(* Logix 5000 project; controller R400_500_XLS vendor 1 type 14 code 216 rev 31.11; software revision 31.01 *)

TASK MainTask (continuous, watchdog 500 ms) : MainProgram

MODULES
   Local : vendor 1 type 14 code 216 (5069 0, rev 31.11)
        LabWasher2:6:O.0   // Audible Alarm/Red Status Light/Alarm Signal Relay
        LabWasher2:6:O.1   // Dry Contact For Cycle Completed or External Pure Water valve
        LabWasher2:6:O.2   // Dry contact For Alarm
        LabWasher2:6:O.3   // Interior Light
        LabWasher2:6:O.4   // Transfer Valve (Normally Open Valve)
        LabWasher2:6:O.5   // Cycle Status Pilot Light
        LabWasher2:6:O.6   // Condensate Return CoolDown water valve
        LabWasher2:6:O.7   // Not Used
        LabWasher2:7:O.0   // Load door close pilot valve
        LabWasher2:7:O.1   // Load door open pilot valve
        LabWasher2:7:O.2   // Unload door close pilot valve
        LabWasher2:7:O.3   // Unload door open pilot valve
        LabWasher2:7:O.4   // Pump low speed
        LabWasher2:7:O.5   // Pump high speed
        LabWasher2:7:O.6   // Hot water sump fill valve
        LabWasher2:7:O.7   // Sump drain valve (Normally open valve)
        LabWasher2:8:O.0   // Vapor removal fan / Drying fan
        LabWasher2:8:O.1   // Sump steam valve/ Electrical Heater
        LabWasher2:8:O.2   // Pure water sump/ Tank fill valve
        LabWasher2:8:O.3   // Drain cool down water valve
        LabWasher2:8:O.4   // Cold water sump fill valve
        LabWasher2:8:O.5   // PWT Steam Valve / Electric Heater
        LabWasher2:8:O.6   // Heat recovery tank drian valve
        LabWasher2:8:O.7   // Pure water tank outlet valve
        LabWasher2:9:O.0   // Drying heating elements
        LabWasher2:9:O.2   // Condenser high flow cold water valve
        LabWasher2:9:O.3   // Condenser low flow cold water valve
        LabWasher2:9:O.4   // Chemical pump #1
        LabWasher2:9:O.5   // Chemical pump #2
        LabWasher2:9:O.6   // Chemical pump #3
        LabWasher2:9:O.7   // Chemical pump #4
        LabWasher2:2:I.0   // Chemical Pump 1 level switch
        LabWasher2:2:I.1   // Chemical Pump #2 level switch
        LabWasher2:2:I.2   // Chemical Pump #3 level switch
        LabWasher2:2:I.3   // Chemical Pump #4 level switch
        LabWasher2:2:I.4   // Pure water tank level switch
        LabWasher2:2:I.5   // Pure water tank safety level switch
        LabWasher2:1:I.0   // Motor overload
        LabWasher2:1:I.1   // MCR input
        LabWasher2:1:I.2   // Load door obstruction switch
        LabWasher2:1:I.3   // Load door close
        LabWasher2:1:I.4   // Sump low level switch
        LabWasher2:1:I.5   // Sump low level switch
        LabWasher2:1:I.6   // Sump safety level switch
        LabWasher2:1:I.7   // Shelf switch
        LabWasher2:3:I.0   // Unload door obstruction switch
        LabWasher2:3:I.1   // Unload door close
        LabWasher2:3:I.2   // Door Open button Unload side
        LabWasher2:3:I.3   // Door Close/ Sielnce button Unload Side
      Serial : vendor 1 type 12 code 320 (5069 1, rev 1.11, StandardDataDriven RPI 80 ms)
      LabWasher2 : 1734-AENT (Ethernet 192.168.1.2, rev 3.4, Output RPI 20 ms)
         IO11 : 1734-IB8 (PointIO 1, rev 3.1)
         IO22 : 1734-IB8 (PointIO 2, rev 3.1)
         IO33 : 1734-IR2 (PointIO 4, rev 3.1, Input RPI 80 ms)
         IO77 : 1734-IR2 (PointIO 5, rev 3.1, Input RPI 80 ms)
         IO66 : 1734-IB8 (PointIO 3, rev 3.1)
         IO99 : 1734-OB8 (PointIO 9, rev 3.1)
         IO88 : 1734-OB8 (PointIO 8, rev 3.1)
         IO44 : 1734-OB8 (PointIO 6, rev 3.1)
         IO55 : 1734-OB8 (PointIO 7, rev 3.1)
      LabWasher : 1734-AENT (Ethernet 192.168.1.4, rev 3.4, Output RPI 20 ms)   // Chamber inputs/outputs remote module
         IO2 : 1734-IB8 (PointIO 2, rev 3.1, Input RPI 20 ms)   // Digital inputs
              LabWasher:2:I.Data.0   // Chemical Pump #1 level switch
              LabWasher:2:I.Data.1   // Chemical Pump #2 level switch
              LabWasher:2:I.Data.2   // Chemical Pump #3 level switch
              LabWasher:2:I.Data.3   // Chemical Pump #4 level switch
              LabWasher:2:I.Data.4   // Pure water tank level switch
              LabWasher:2:I.Data.5   // Pure water tank safety level switch
              LabWasher:2:I.Data.6   // Pure Water Filling Authorization Signal
         IO3 : 1734-IR2 (PointIO 4, rev 3.1, Input RPI 80 ms)   // Analog input
              LabWasher:4:I.Ch0Data   // Sump RTD
              LabWasher:4:I.Ch1Data   // Drying RTD
              LabWasher:4:I.Ch0Fault   // Sump RTD channel Fault bit
              LabWasher:4:I.Ch1Fault   // Dry RTD channel Fault bit
         IO7 : 1734-IR2 (PointIO 5, rev 3.1, Input RPI 80 ms)   // RTD inputs
              LabWasher:5:I.Ch0Data   // Pure Water Tank RTD
              LabWasher:5:I.Ch1Data   // Not Used
              LabWasher:5:I.Ch0Fault   // Pure Water Tank RTD channel Fault bit
         IO10 : 1734-IE4C (PointIO 10, rev 3.1, Input RPI 80 ms)   // Analog inputs
              LabWasher:10:I.Ch0Data   // Chemical water conductivity
              LabWasher:10:I.Ch1Data   // Final rinse water conductivity
              LabWasher:10:I.Ch2Data   // Recirculation pump pressure
              LabWasher:10:I.Ch3Data   // Not Used
              LabWasher:10:I.Ch0Fault   // Chemical conductivity channel Fault bit
              LabWasher:10:I.Ch1Fault   // Final rinse conductivity channel Fault bit
              LabWasher:10:I.Ch2Fault   // Pressure Transmitter analog channel Fault bit
         IO6 : 1734-IB8 (PointIO 3, rev 3.1, Input RPI 20 ms)   // Digital input
              LabWasher:3:I.Data.0   // Unload door obstruction switch
              LabWasher:3:I.Data.1   // Unload door close
              LabWasher:3:I.Data.2   // Door Open button Unload side
              LabWasher:3:I.Data.3   // Door Close/ Sielnce button Unload Side
              LabWasher:3:I.Data.4   // Not Used
              LabWasher:3:I.Data.5   // Not Used
              LabWasher:3:I.Data.6   // Not Used
              LabWasher:3:I.Data.7   // Not Used
         IO1 : 1734-IB8 (PointIO 1, rev 3.1, Input RPI 20 ms)   // Digital inputs
              LabWasher:1:I.Data.0   // Motor overload
              LabWasher:1:I.Data.1   // MCR input
              LabWasher:1:I.Data.2   // Load door obstruction switch
              LabWasher:1:I.Data.3   // Load door close
              LabWasher:1:I.Data.4   // Sump low level switch
              LabWasher:1:I.Data.5   // Sump high level switch
              LabWasher:1:I.Data.6   // Sump safety level switch
              LabWasher:1:I.Data.7   // Shelf switch
         IO8 : 1734-OB8 (PointIO 8, rev 3.1, Output RPI 20 ms)   // Digital outputs
              LabWasher:8:O.Data.0   // Vapor removal fan / Drying fan
              LabWasher:8:O.Data.1   // Sump steam valve/ Electrical Heater
              LabWasher:8:O.Data.2   // Pure water sump/ Tank fill valve
              LabWasher:8:O.Data.3   // Drain cool down water valve
              LabWasher:8:O.Data.4   // Cold water sump fill valve
              LabWasher:8:O.Data.5   // PWT Steam Valve / Electric Heater
              LabWasher:8:O.Data.6   // Heat recovery tank drian valve
              LabWasher:8:O.Data.7   // Pure water tank outlet valve
         IO4 : 1734-OB8 (PointIO 6, rev 3.1, Output RPI 20 ms)   // Digital output
              LabWasher:6:O.Data.0   // Audible Alarm/Red Status Light/Alarm Signal Relay
              LabWasher:6:O.Data.1   // Dry Contact For Cycle Completed or External Pure Water valve
              LabWasher:6:O.Data.2   // Dry contact For Alarm
              LabWasher:6:O.Data.3   // Interior Light
              LabWasher:6:O.Data.4   // Transfer Valve (Normally Open Valve)
              LabWasher:6:O.Data.5   // Cycle Status Pilot Light
              LabWasher:6:O.Data.6   // Condensate Return CoolDown water valve
              LabWasher:6:O.Data.7   // Not Used
         IO5 : 1734-OB8 (PointIO 7, rev 3.1, Output RPI 20 ms)   // Digital output
              LabWasher:7:O.Data.0   // Load door close pilot valve
              LabWasher:7:O.Data.1   // Load door open pilot valve
              LabWasher:7:O.Data.2   // Unload door close pilot valve
              LabWasher:7:O.Data.3   // Unload door open pilot valve
              LabWasher:7:O.Data.4   // Pump low speed
              LabWasher:7:O.Data.5   // Pump high speed
              LabWasher:7:O.Data.6   // Hot water sump fill valve
              LabWasher:7:O.Data.7   // Sump drain valve (Normally open valve)
         IO9 : 1734-OB8 (PointIO 9, rev 3.1, Output RPI 20 ms)   // Digital outputs
              LabWasher:9:O.Data.0   // Drying heating elements
              LabWasher:9:O.Data.1   // Drying Isolation Valve (Normally Closed Valve)
              LabWasher:9:O.Data.2   // Condenser high flow cold water valve
              LabWasher:9:O.Data.3   // Condenser low flow cold water valve
              LabWasher:9:O.Data.4   // Chemical pump #1
              LabWasher:9:O.Data.5   // Chemical pump #2
              LabWasher:9:O.Data.6   // Chemical pump #3
              LabWasher:9:O.Data.7   // Chemical pump #4
END_MODULES

TYPE FaultRecord :
STRUCT
   TimeLow : DINT;   // Lower 32 bits of the fault timestamp value
   TimeHigh : DINT;   // Upper 32 bits of the fault timestamp value
   Type : INT;   // Fault type (program, I/O, etc.)
   Code : INT;   // Unique code for the fault
   Info : DINT[8];   // Fault specific information
END_STRUCT
END_TYPE

TYPE Hrdwre :
STRUCT
   Model : BOOL;   // Reliance Mdl 400 = 0 500 = 1
   NbDoors : BOOL;   // Single = 0 Double =1
   PreWtrTnk : BOOL;   // Pure Water Tank Option 1= Yes
   HtRcvryTnk : BOOL;   // Heat Recovery Tank Option 1= Yes
   Dry : BOOL;   // Drying Option
   ElectricUnit : BOOL;   // Electric Heated Unit 1= Electric
   CoolDown : BOOL;   // Drain Cooldown Option 1= Yes 0 = No
   NbChmPmp : SINT;   // 2, 3 or 4 chemical pumps
   Condenser : BOOL;   // With Condenser = 1
   CWInlet : BOOL;   // With Cold Water Inlet Option = 1
   MonitorPressure : BOOL;   // 0 = No pressure monitoring, 1 = Pressure monitoring
   MonitorCond : BOOL;   // 0 = No conductivity monitoring, 1 = Conductivity monitoring
   CondensateReturn : BOOL;   // Condensate Return Option
   Printer : BOOL;   // 1 = Printer option present
   EmailNotification : BOOL;   // 1= Email & SMS Notification Enable (PLC & HMI)
   AuditTrail : BOOL;   // 1 = With Audit Trail
   BatchReport : BOOL;   // 1 = With Batch Report
   CycleValidation : BOOL;   // 1 = With Cycle Validation
   ElectronicSignature : BOOL;   // 1 = With Electronic Signature
END_STRUCT
END_TYPE

TYPE List :
STRUCT
   Value : DINT;
   Ind : DINT;
   Rmte : BOOL;
   Enter : BOOL;
END_STRUCT
END_TYPE

TYPE NameLocation :
STRUCT
   Pos1 : STRING;   // Cycle Name Position 1
   Pos2 : STRING;   // Cycle Name Position 2
   Pos3 : STRING;   // Cycle Name Position 3
   Pos4 : STRING;   // Cycle Name Position 4
   Pos5 : STRING;   // Cycle Name Position 5
   Pos6 : STRING;   // Cycle Name Position 6
   Pos7 : STRING;   // Cycle Name Position 7
   Pos8 : STRING;   // Cycle Name Position 8
   Pos9 : STRING;   // Cycle Name Position 9
   Pos10 : STRING;   // Cycle Name Position 10
   Pos11 : STRING;   // Cycle Name Position 11
   Current : STRING;   // Name of the current cycle
END_STRUCT
END_TYPE

TYPE UDT_AuditTrail :
STRUCT
   bCapacityHighWarning : BOOL;   // Capacity High Warning
   bCapacityHighHighWarning : BOOL;   // Capacity High High Warning
   bRemoteClearAuditHistory : BOOL;   // Remote Clear Audit History
END_STRUCT
END_TYPE

TYPE UDT_CHEM_PUMP :   // Flow rate of the chemical pump 4
STRUCT
   FlowRate : DINT;   // Flow rate of the chemical pump 1
END_STRUCT
END_TYPE

TYPE UDT_CSVDataLog :   // CSV Data Log
STRUCT
   sFileLocation : STRING;   // File Location
   bTrigger : BOOL;   // Trigger
   sString01 : STRING;   // String #1
   bHandshake : BOOL;   // Handshake
END_STRUCT
END_TYPE

TYPE UDT_CSVExport :   // CSV Export
STRUCT
   bExportTrigger : BOOL;   // Trigger
   sFileLabel : STRING;   // File Name
   iStatusCode : DINT;   // Status Code
   sStatusMessage : STRING;   // Status Message
   bExportTriggerUnloadSideHMI : BOOL;   // Trigger for a Unload Side HMI
END_STRUCT
END_TYPE

TYPE UDT_CYCLE :   // UDT CYCLE
STRUCT
   PW : UDT_PW[4];   // Pre-Wash Treatments
   WSH : UDT_WASH[5];   // Wash Treatments
   RINSE : UDT_RINSE[4];   // Rinse treatments
   FRINSE : UDT_FRINSE;   // F rinse treatments
   DRY : UDT_DRY;   // Dry Treatment
   Lock : BOOL;   // Cycle permission 1= Cycle is unlocked
   AutoWtrLevel : BOOL;   // Auto Water Level 0= Auto 1 = High Level
   AutoSpeed : BOOL;   // Auto Speed 0 = Auto 1= Low
END_STRUCT
END_TYPE

TYPE UDT_CYCLE_SEQUENCE :
STRUCT
   InitialStep : BOOL;
   PreWash1Start : BOOL;
   PreWash1End : BOOL;
   PreWash2Start : BOOL;
   PreWash2End : BOOL;
   PreWash3Start : BOOL;
   PreWash3End : BOOL;
   PreWash4Start : BOOL;
   PreWash4End : BOOL;
   Wash1Start : BOOL;
   Wash1End : BOOL;
   Wash2Start : BOOL;
   Wash2End : BOOL;
   Wash3Start : BOOL;
   Wash3End : BOOL;
   Wash4Start : BOOL;
   Wash4End : BOOL;
   Wash5Start : BOOL;
   Wash5End : BOOL;
   Rinse1Start : BOOL;
   Rinse1End : BOOL;
   Rinse2Start : BOOL;
   Rinse2End : BOOL;
   Rinse3Start : BOOL;
   Rinse3End : BOOL;
   Rinse4Start : BOOL;
   Rinse4End : BOOL;
   FinalRinseStart : BOOL;
   FinalRinseEnd : BOOL;
   DryingStart : BOOL;
   DryingEnd : BOOL;
   VentingStart : BOOL;
   VentingEnd : BOOL;
END_STRUCT
END_TYPE

TYPE UDT_CYCLE_USAGE :   // Cycle Usage
STRUCT
   UserName : STRING;   // Name of the user
   CycleStartedCount : DINT;   // Count the Number Of time a user start a Cycle
END_STRUCT
END_TYPE

TYPE UDT_DRY :   // Data Type of a Drying.
STRUCT
   Trt : INT;   // Treatment Number 18 = Drying
   Mode : INT;   // Drying Mode 0 = Smart 1= Standard
   Tmin : INT;   // Drying time in Minute
   Tsec : INT;   // Drying time in Second
   HiLowTemp : BOOL;   // 1= High 115.6 C 0 = 82.2 C
   HeatSensitive : BOOL;   // 0 = Regular 1= Heat Sensitive
END_STRUCT
END_TYPE

TYPE UDT_FRINSE :   // Data Type of a Final Rinse.
STRUCT
   Trt : INT;   // Final Rinse Treatment Number
   Prt : INT;   // Final Rinse Water Port
   Heat : BOOL;   // Final Rinse Heated =1, Non-Heated = 0
   Tmp : REAL;   // Final Rinse Temperature
   Tmin : INT;   // Final Rinse Time in Minute
   Tsec : INT;   // Final Rinse Time in Second
   Type : INT;   // Final Rinse Type
   Nb : INT;   // Number of Final Rinses
   MnNb : INT;   // Minimum number of Rinses
   CondSP : REAL;   // Final Rinse Conductivity Set Point
   Recirc : BOOL;   // recirculated final rinse 1 = Yes
   Drn : BOOL;   // 0 = Water Saved 1= Water Drained
END_STRUCT
END_TYPE

TYPE UDT_NUMERIC_INPUT :   // Data type reprensenting the numeric input control in FT View
STRUCT
   value : DINT;   // Value of the numeric input
   caption : DINT;   // Value displayed on the numeric screen
   enter : BOOL;   // Set when the enter key is pressed
   hds : BOOL;   // Reset the enter connection
END_STRUCT
END_TYPE

TYPE UDT_NUMERIC_INPUT_REAL :   // Handskake
STRUCT
   value : REAL;   // Write Tag
   caption : REAL;   // Read tag
   enter : BOOL;   // Enter
   hds : BOOL;   // Handskake
END_STRUCT
END_TYPE

TYPE UDT_PORT_HANDSHAKE_FROM_SCADA :
STRUCT
   bFillingAuthorizationSignal : BOOL;   // Pure Water Filling Authroization Signal
END_STRUCT
END_TYPE

TYPE UDT_PORT_HANDSHAKE_TO_SCADA :   // Pure Water Handshake to SCADA
STRUCT
   bFillRequest : BOOL;   // Pure Water Filling Request
   bLoopValve : BOOL;   // Pure Water Loop Valve
END_STRUCT
END_TYPE

TYPE UDT_PW :   // UDT PRE-WASH
STRUCT
   TrtNo : DINT;   // Treatment Number
   Wprt : DINT;   // Water Port 1= Cold Water 2= Hot Water
   Heat : BOOL;   // 1 = Heated
   Tmp : REAL;   // TempSp
   Tmin : INT;   // Temps Min
   Tsec : INT;   // Temps Sec
END_STRUCT
END_TYPE

TYPE UDT_RINSE :   // UDT RINSE TREATMENT
STRUCT
   TrtNo : DINT;   // Treatment Number
   Wprt : DINT;   // Water Port 1= Cold Water 2= Hot Water
   Heat : BOOL;   // 1 = Heated
   Tmp : REAL;   // TempSp
   Tmin : INT;   // Temps Min
   Tsec : INT;   // Temps Sec
END_STRUCT
END_TYPE

TYPE UDT_SCALE :   // Data type used for scaling the analog inputs
STRUCT
   InputMin : DINT;   // Minimum Raw Data
   InputMax : DINT;   // Maximum Raw Data
   ScaledMin : REAL;   // Minimum Scaled Data
   ScaledMax : REAL;   // Maximum Scaled Data
   DfInputMin : DINT;   // Default Minimum Raw Data
   DfInputMax : DINT;   // Default Maximum raw Data
   DfScaledMin : DINT;   // Default Minimum Scaled Data
   DfScaledMax : DINT;   // Default Maximum Scaled Data
   Input : DINT;   // Raw Input Value
   Output : REAL;   // Scaled Output
END_STRUCT
END_TYPE

TYPE UDT_SELECTOR :   // This data type represent the HMI piloted list selector
STRUCT
   Value : INT;   // Position of the selector
   Indicator : INT;   // Position set by the PLC
   Remote : BOOL;   // Remote control
END_STRUCT
END_TYPE

TYPE UDT_STRING_INPUT :
STRUCT
   Value : STRING;   // String Value
   Caption : STRING;   // String Display
   Enter : BOOL;   // String input Enter Key
   Hds : BOOL;   // String Handshake
END_STRUCT
END_TYPE

TYPE UDT_TCPSetAllConfig :
STRUCT
   IPAddress : DINT;   // IPaddress
   SunbNetMask : DINT;   // Subnet Mask
   Gateway : DINT;   // Gateway IP address
   NameServer1 : DINT;   // Primary DNS Server IP address
   NameServer2 : DINT;   // Secondary DNS Server IP address
   DomainName : SINT[50];
END_STRUCT
END_TYPE

TYPE UDT_WASH :   // UDT Wash treatment
STRUCT
   TrtNo : DINT;   // Treatment Number
   Wprt : DINT;   // Water Port 1= Cold Water 2= Hot Water
   Heat : BOOL;   // 1 = Heated
   Tmp : REAL;   // TempSp
   Tmin : INT;   // Temps Min
   Tsec : INT;   // Temps Sec
   ChemUsed_1 : INT;   // Chemi 1st Injection
   ChemUsed_2 : INT;   // Chem 2nd Injection
   InjType_1 : BOOL;   // Inj Type 1st Injection
   InjType_2 : BOOL;   // Inj. Type 2nd Injection
   ChemVol_1 : REAL;   // Chem Volume 1st Injection
   ChemVol_2 : REAL;   // Chem Volume 2nd injection
   CondSp_1 : REAL;   // Cond Sp 1st Injection
   CondSp_2 : REAL;   // Cond Sp 2nd Injection
END_STRUCT
END_TYPE

ADD_ON_INSTRUCTION Doors   (* revision 1.0 *)
VAR_IN_OUT
   Displayed : DINT; {required}
END_VAR
VAR_INPUT
   Obstruction : BOOL; {required}
   Closed : BOOL; {required}
END_VAR
VAR_IN_OUT
   ClosePressed : BOOL; {required}
END_VAR
VAR_INPUT
   PreviousScreen : DINT; {required}
END_VAR
VAR_IN_OUT
   OpenPressed : BOOL; {required}
END_VAR
VAR_OUTPUT
   Open : BOOL; {access Read Only, required}
   Closing : BOOL; {access Read Only, required}
END_VAR
VAR_IN_OUT
   StopPressed : BOOL; {required}
   Msg1 : INT; {required}
END_VAR
VAR_INPUT
   ServiceMode : BOOL; {required}
   AutoClosing : BOOL; {required}
   Delay12S : DINT; {required}
   Delay1250ms : DINT; {required}
END_VAR
VAR_OUTPUT
   Step15 : BOOL; {access Read Only, required}   // Maintain close
   Step12 : BOOL; {access Read Only, required}   // Maintain open
END_VAR
VAR_INPUT
   MsgOpening : INT; {required}
   MsgClosing : INT; {required}
END_VAR
VAR_OUTPUT
   Step17 : BOOL; {access Read Only, required}   // Alarm Obstruction
   Step16 : BOOL; {access Read Only, required}   // Alarm door not close
   Step13 : BOOL; {access Read Only, required}   // Alarm door not open
   Step11 : BOOL; {access Read Only, required}   // Opening
   Step14 : BOOL; {access Read Only, required}   // Closing
END_VAR
VAR_INPUT
   CurrentScreen : DINT; {required}
END_VAR
VAR
   ONS1 : BOOL;
   Doors : BOOL;
   ONS2 : BOOL;
   ONS3 : BOOL;
   ONS4 : BOOL;
   ONS5 : BOOL;
   s108 : DINT := 108;   // Screen 108
   Ons6 : BOOL;
   Ons7 : BOOL;
   OpeningDelay : TIMER := (PRE := 12000);
   ClosingDelay : TIMER;
   OpenDelayAlarm : TIMER;
   Step10 : BOOL := 1;   // Waiting
   RequestScreen : DINT;   // Request Screen When Available
END_VAR

ROUTINE Logic   (* ladder *)
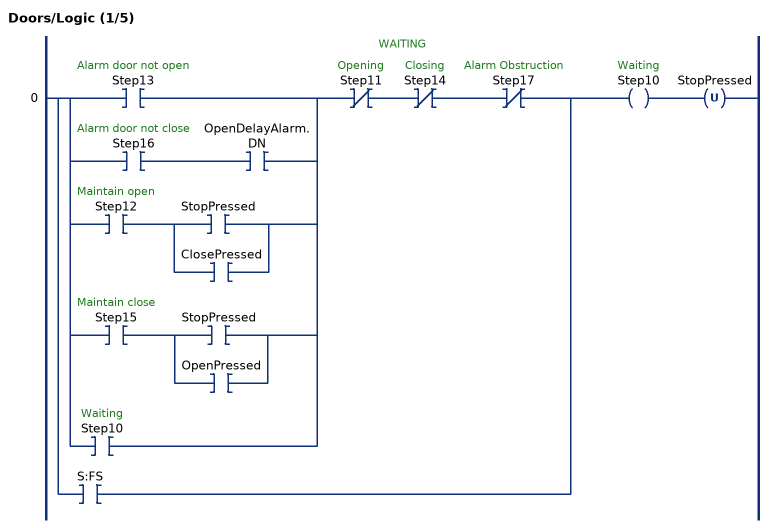
   // WAITING
   0: [[XIC(Step13) ,XIC(Step16) XIC(OpenDelayAlarm.DN) ,XIC(Step12) [XIC(StopPressed) ,XIC(ClosePressed) ] ,XIC(Step15) [XIC(StopPressed) ,XIC(OpenPressed) ] ,XIC(Step10) ] XIO(Step11) XIO(Step14) XIO(Step17) ,XIC(S:FS) ]OTE(Step10)OTU(StopPressed);
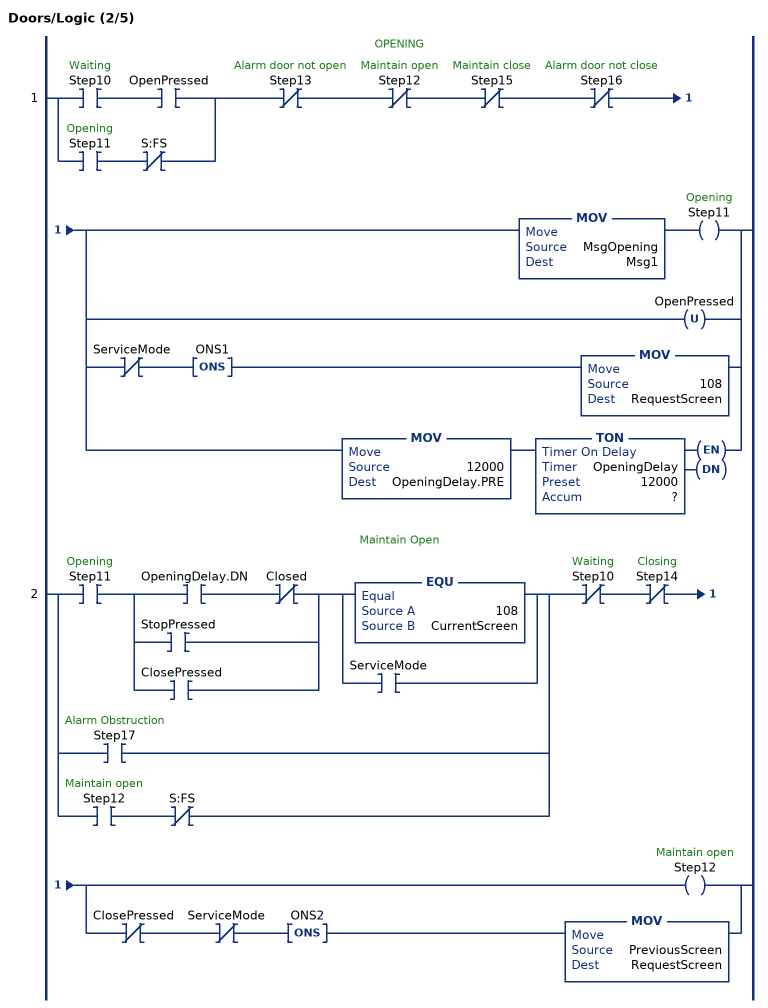
   // OPENING
   1: [XIC(Step10) XIC(OpenPressed) ,XIC(Step11) XIO(S:FS) ]XIO(Step13)XIO(Step12)XIO(Step15)XIO(Step16)[MOV(MsgOpening,Msg1) OTE(Step11) ,OTU(OpenPressed) ,XIO(ServiceMode) ONS(ONS1) MOV(108,RequestScreen) ,MOV(12000,OpeningDelay.PRE) TON(OpeningDelay,?,?) ];
   // Maintain Open
   2: [[XIC(Step11) [XIC(OpeningDelay.DN) XIO(Closed) ,XIC(StopPressed) ,XIC(ClosePressed) ] [EQU(108,CurrentScreen) ,XIC(ServiceMode) ] ,XIC(Step17) ] ,XIC(Step12) XIO(S:FS) ]XIO(Step10)XIO(Step14)[OTE(Step12) ,XIO(ClosePressed) XIO(ServiceMode) ONS(ONS2) MOV(PreviousScreen,RequestScreen) ];
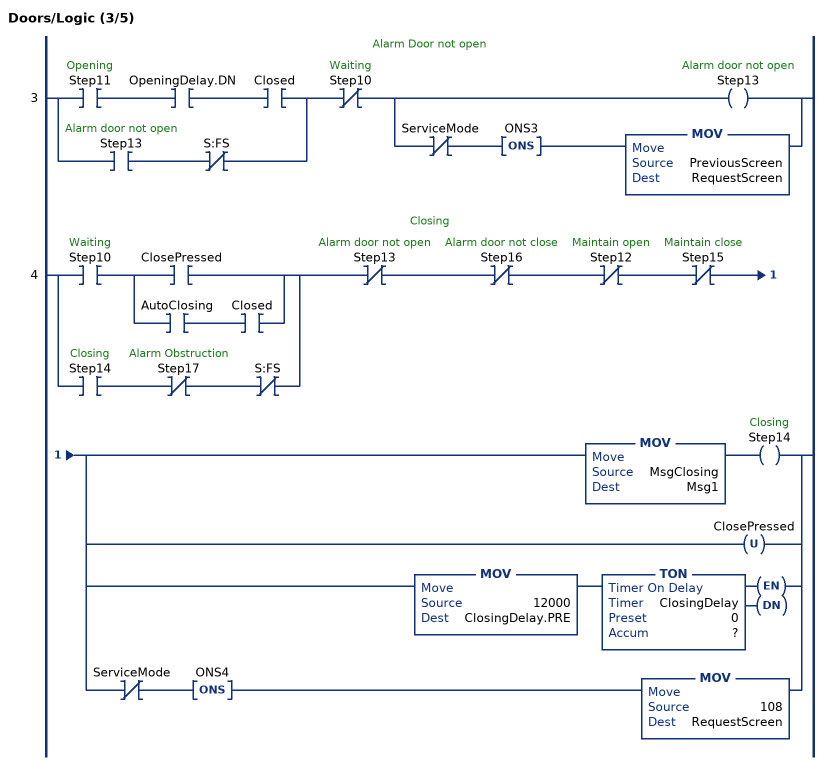
   // Alarm Door not open
   3: [XIC(Step11) XIC(OpeningDelay.DN) XIC(Closed) ,XIC(Step13) XIO(S:FS) ]XIO(Step10)[OTE(Step13) ,XIO(ServiceMode) ONS(ONS3) MOV(PreviousScreen,RequestScreen) ];
   // Closing
   4: [XIC(Step10) [XIC(ClosePressed) ,XIC(AutoClosing) XIC(Closed) ] ,XIC(Step14) XIO(Step17) XIO(S:FS) ]XIO(Step13)XIO(Step16)XIO(Step12)XIO(Step15)[MOV(MsgClosing,Msg1) OTE(Step14) ,OTU(ClosePressed) ,MOV(12000,ClosingDelay.PRE) TON(ClosingDelay,?,?) ,XIO(ServiceMode) ONS(ONS4) MOV(108,RequestScreen) ];
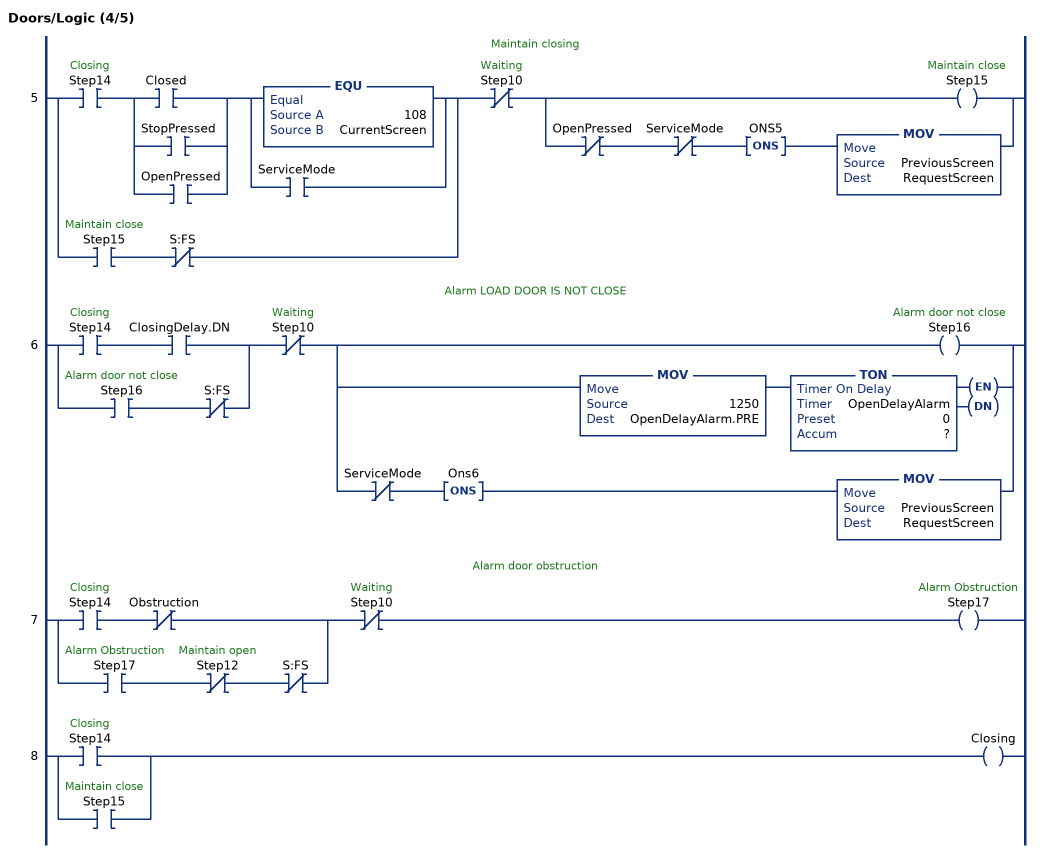
   // Maintain closing
   5: [XIC(Step14) [XIC(Closed) ,XIC(StopPressed) ,XIC(OpenPressed) ] [EQU(108,CurrentScreen) ,XIC(ServiceMode) ] ,XIC(Step15) XIO(S:FS) ]XIO(Step10)[OTE(Step15) ,XIO(OpenPressed) XIO(ServiceMode) ONS(ONS5) MOV(PreviousScreen,RequestScreen) ];
   // Alarm LOAD DOOR IS NOT CLOSE
   6: [XIC(Step14) XIC(ClosingDelay.DN) ,XIC(Step16) XIO(S:FS) ]XIO(Step10)[OTE(Step16) ,MOV(1250,OpenDelayAlarm.PRE) TON(OpenDelayAlarm,?,?) ,XIO(ServiceMode) ONS(Ons6) MOV(PreviousScreen,RequestScreen) ];
   // Alarm door obstruction
   7: [XIC(Step14) XIO(Obstruction) ,XIC(Step17) XIO(Step12) XIO(S:FS) ]XIO(Step10)OTE(Step17);
   8: [XIC(Step14) ,XIC(Step15) ]OTE(Closing);
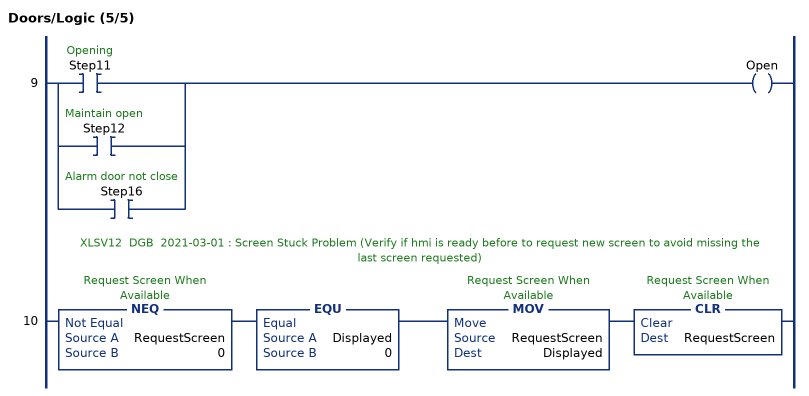
   9: [XIC(Step11) ,XIC(Step12) ,XIC(Step16) ]OTE(Open);
   // XLSV12  DGB  2021-03-01 : Screen Stuck Problem (Verify if hmi is ready before to request new screen to avoid missing the last screen requested)
   10: NEQ(RequestScreen,0)EQU(Displayed,0)MOV(RequestScreen,Displayed)CLR(RequestScreen);
END_ROUTINE
END_ADD_ON_INSTRUCTION

VAR_GLOBAL   (* controller tags *)
   abCycleDataToSCADA : BOOL[32];
   abInputToSCADA : BOOL[32] := ([1] := 1, [2] := 1, [3] := 1, [6] := 1, [7] := 1, [8] := 1, [9] := 1, [13] := 1, [14] := 1);
   abOutputToSCADA : BOOL[32] := ([2] := 1, [3] := 1, [8] := 1, [15] := 1, [23] := 1);
   ActualDay : DINT := 9716;
   aiCycleDataToSCADA : INT[16] := ([2] := 14, [3] := 16, [4] := 52, [6] := 24, [7] := 49, [8] := 60);
   AlarmAck : INT;   // Alarm acknowledgement from the HMI
   AlarmMsg : STRING := 'MAINTENANCE DUE';   // Message of the alarm from the HMI Do not delete this tag
   AlarmTrigger : INT;   // Triggers the alarm screen if different of 0
   arAnalogInputToSCADA : REAL[8] := ([0] := 0.1, [1] := 34.34375, [2] := 32.122498, [4] := 21.7, [5] := 22.798864, [6] := 21.9);
   arCycleDataToSCADA : REAL[8] := ([2] := 1.4172212, [3] := 11.417221);
   bAcceptRejectRecorded : BOOL := 1;   // Cycle Accept/Reject Recorded By User
   BatteryLowWarning : BOOL;
   bAuditTrailExportButton : BOOL;
   bCSVExportHandshake : BOOL;
   bCycleOrAbortInProcess : BOOL;
   bFactoryReset : BOOL;
   bFactoryResetCompleted : BOOL;
   bHMICycleAccepted : BOOL;   // HMI - Button Cycle Accepted
   bHMICycleRejected : BOOL;   // HMI - Button Cycle Rejected
   bInibitAutologout : BOOL := 1;   // Cancel AutoLogout
   bNewStringDetected : BOOL;
   BoilingValue : REAL := 100.03;
   bONSAuditExportTrigger : BOOL;
   bONSAuditTrailAlarm : BOOL;
   bONSAuditTrailEndOfCycle : BOOL := 1;
   bONSBatchReportFileLocation : BOOL;
   bONSCycleAccepted : BOOL;
   bONSCycleRejected : BOOL;
   bONSFactoryReset : BOOL;
   bONSManualFileTransfer : BOOL;
   bONSSerialModuleResetInhibit : BOOL := 1;
   bONSSerialModuleSetInhibit : BOOL;
   bPureWaterFillingAuthorization : BOOL := 1;   // Pure Water Filling Authorization Signal
   bPushButtonTransferFilesFromSDToUSB : BOOL;
   bResetHardwareOptions : BOOL;
   bResetModulesConfiguration : BOOL;
   bResetSystemOptions : BOOL;
   bSerialModuleConfigureInhibit : BOOL;   // Configure if Serial Card is Inhibited or not
   bTransferFilesFromSDToUSB : BOOL;
   bTransferFilesFromSDToUSBHandshakeLoad : BOOL;
   CalibCounter : SINT;
   Cfg_10_Modules : BOOL := 1;   // Chassis is configured 10 slots
   Cfg_11_Modules : BOOL;
   CfgChem : SINT;
   CfgChem2 : SINT;
   CfgConc : REAL;
   CfgConc2 : REAL;
   CfgCondSp : REAL;
   CfgInjType : SINT;
   cfgPrewashHeated : SINT;
   cfgPrewashMin : SINT;
   cfgPrewashSec : DINT;
   CfgPrewashTempSp : REAL := 65.6;
   cfgPrewashWport : SINT := 2;
   cfgRinseHeated : SINT;
   cfgRinseMin : SINT;
   cfgRinseSec : SINT;
   CfgRinseTempSp : REAL := 80.0;
   cfgRinseWport : SINT := 2;
   CfgWshHeated : SINT := 1;
   CfgWshInjRateImperial : REAL := 0.5;   // Wash Injection Rate - Oz / Gal
   CfgWshInjRateMetric : REAL := 1.0;   // Wash Injection Rate - mL / L
   CfgWshMin : SINT;
   CfgWshSec : SINT;
   CfgWshTempSp : REAL := 70.0;
   cfgWshWport : SINT := 2;
   ChangeLanguage : BOOL;   // Tag Changed By HMI To Start Printout Message Translation
   Chassis_Size_Ret : DINT[3];
   ChemConcUnit : BOOL := 1;   // 0 = mL/L; 1 = oz/gal
   ChemCond : REAL := 0.1;
   ChemicalName : STRING[9] := ([1] := 'CIP 100', [2] := 'CIP 200', [3] := 'N/A', [4] := 'N/A', [6] := 'N/A', [7] := 'Pump 3', [8] := 'Pump 4');   // Used by HMI
   ChemPumpSelector : UDT_SELECTOR[2];   // Chemical pump calibration selector
   COOLING_PHASE_TIME : DINT := 120000;   // Time of the cooling phase when time based drying
   CR2Mode : SINT := 1;   // 0= Cycle complete dry contact 1= External pure water valve
   Ctrlr_Status : DINT := 4448;
        .13   // Compact Logix Key Status 1= Key in Rmte or Prog Pos. 0 = Key in Run Pos.
   Current_Screen : DINT := 99;
   CurrentUser : STRING := 'service';   // Current User
   CycleCounter : DINT := 60;
   CycleName : STRING[12] := ([0] := 'CYCLE 1', [1] := 'HEAVY', [2] := 'COUPONS', [3] := 'DRY', [4] := 'BINS', [5] := 'NODET 6', [6] := 'LUKE 0', [7] := 'CYCLE 8', [8] := 'STERIS', [9] := 'CYCLE 10', [10] := 'STERIS', [11] := 'STERIS');
        [11]   // Cycle Name Buffer
   CycleNameDefault : STRING[12] := ([0] := 'EXTRACare', [1] := 'ENVIROCare', [2] := 'PLASTIC', [3] := 'STANDARD', [4] := 'RINSECare', [5] := 'DESCALER', [6] := 'CYCLE 7', [7] := 'CYCLE 8', [8] := 'CYCLE 9', [9] := 'CYCLE 10', [10] := 'CYCLE 11');
   CyclePtr : DINT := 8;   // Cycle Pointeur
   CycleUsage : UDT_CYCLE_USAGE[50] := ([0].UserName := 'service', [0].CycleStartedCount := 60, [1].UserName := 'User 03', [1].CycleStartedCount := 1, [2].UserName := '-', [3].UserName := '-', [4].UserName := '-', [5].UserName := '-', [6].UserName := '-', [7].UserName := '-', [8].UserName := '-', [9].UserName := '-', [10].UserName := '-', [11].UserName := '-', [12].UserName := '-', [13].UserName := '-', [14].UserName := '-', [15].UserName := '-', [16].UserName := '-', [17].UserName := '-', [18].UserName := '-', [19].UserName := '-', [20].UserName := '-', [21].UserName := '-', [22].UserName := '-', [23].UserName := '-', [24].UserName := '-', [25].UserName := '-', [26].UserName := '-', [27].UserName := '-', [28].UserName := '-', [29].UserName := '-', [30].UserName := '-', [31].UserName := '-', [32].UserName := '-', [33].UserName := '-', [34].UserName := '-', [35].UserName := '-', [36].UserName := '-', [37].UserName := '-', [38].UserName := '-', [39].UserName := '-', [40].UserName := '-', [41].UserName := '-', [42].UserName := '-', [43].UserName := '-', [44].UserName := '-', [45].UserName := '-', [46].UserName := '-', [47].UserName := '-', [48].UserName := '-', [49].UserName := '-');
   CycleUsageListSelectedIndex : DINT;   // Current index selected in CycleUsage list
   CycleUsagePrint : BOOL;   // Print Cycle Usage
   CycleUsageResetAllValues : BOOL;   // Reset All Cycle Usage of all user
   CycleUsageResetDate : DINT[7] := ([0] := 2022, [1] := 5, [2] := 13, [3] := 13, [4] := 42, [5] := 56, [6] := 51848);
   CycleUsageResetSelectedUser : BOOL;   // Reset Cycle Usage for the selected user
   DateFormat : SINT := 1;   // 0: M-D-Y 1: D-M-Y 2: Y-M-D
   DateTime : DINT[7] := ([0] := 2026, [1] := 8, [2] := 17, [3] := 11, [4] := 1, [5] := 28, [6] := 858318);
        [0]   // PLC Year
        [1]   // PLC Month
        [2]   // PLC Date
        [3]   // PLC Hour
        [4]   // PLC Min
        [5]   // PLC sec.
        [6]   // PLC Microseconds
   DateTimeNew : DINT[7] := ([0] := 2026, [1] := 8, [2] := 13, [3] := 9, [4] := 43, [5] := 47, [6] := 1);
   DISABLE : BOOL;   // Disable bit
   Doors_Check : DINT := 1;
        .0   // Initial Step
        .1   // Yes button has been pressed
        .10   // Door_Check_Step
        .11   // Door_Check_Step
        .12   // Door_Check_Step
        .13   // Door_Check_Step
        .14   // NOT USED
        .15   // Door_Check_Step
        .16   // Test Cancelled
        .17   // Door_Check_Step
        .18   // NOT USED
        .19   // Door_Check_Step
        .2   // No Button Pressed
        .20   // Door_Check_Step
        .21   // Door_Check_Step
        .22   // Door_Check_Step
        .23   // Door_Check_Step
        .24   // Door_Check_Step
        .25   // Door_Check_Step
        .26   // Door_Check_Step
        .27   // Door_Check_Step
        .28   // NOT USED
        .29   // Door_Check_Step
        .3   // Yes Button Pressed
        .30   // Disable Unload Door Open Alarm
        .4   // Door_Check_Step
        .5   // Door_Check_Step
        .6   // Door_Check_Step
        .7   // Door_Check_Step
        .8   // Door_Check_Step
        .9   // Door_Check_Step
   DoorSafetyCheck : BOOL;
   DoorSafetyCheckDay : DINT := 12;
   DoorSafetyCheckMonth : DINT := 8;
   DoorSafetyCheckYear : DINT := 2026;
   DrainExtensionTime : DINT;
   DryTemp : REAL := 22.798864;
   EmailSMSInt : INT[8] := ([6] := 8);   // Email & SMS Notification Integer
        [0]   // Email Command
        [1]   // Email Options
        [1].0   // Email Cycle Started
        [1].1   // Email Cycle Completed
        [1].10   // Email Process Alarms
        [1].2   // Email Cycle Aborted
        [1].3   // Email Cycle Values Changed
        [1].6   // Email Service Mode Entered
        [1].7   // Email Superviser Mode Entered
        [1].8   // Not Used
        [2]   // Email + Text Send Control
        [2].0   // Email ActiveX Trigger
        [2].1   // Email Macro2 Update
        [2].3   // Email ActiveX Handshake
        [2].4   // Email Send Retry
        [2].5   // Email ActiveX Failure Code
        [2].6   // Email ActiveX Failure Code Latch
        [2].7   // Text Macro3 Update
        [3]   // ONS
        [3].0   // ONS used
        [3].1   // ONS used
        [3].10   // ONS used
        [3].15   // Not Used
        [3].2   // ONS used
        [3].3   // ONS used
        [3].4   // ONS used
        [3].5   // ONS used
        [3].6   // ONS used
        [3].7   // ONS used
        [3].8   // Not Used
        [3].9   // DataStore Plus Write Request
        [4]   // Email Retry Counter
        [5]   // PMPack HMI Number
        [6]   // Previous Month
        [7]   // Cell and/or Email Selection
   ENABLE : BOOL := 1;   // Enable bit
   EnaDisPrinter : BOOL := 1;   // Screen 80 Enable/Disable Printer button
   EnDis_LabWasher : DINT := 4;
   EnDis_LabWasher2 : DINT;
   Ethernet_Config_Msg : MESSAGE;
        MessageParameters(ServiceCode := 16#0010, LocalElement := Set_TCP_Config, ...)
   Ethernet_Flash_Write_Msg : MESSAGE;
        MessageParameters(ServiceCode := 16#0010, LocalElement := Set_ConfigControl, ...)
   F8 : REAL[6] := ([0] := 219.0, [1] := 849.0, [2] := 223.0, [3] := 9495.0, [4] := 4000.0, [5] := 12566.0);
        [0]   // Sump RTD
        [1]   // Pure Water Tank RTD
        [2]   // Drying RTD
        [3]   // Final Rinse conductivity
        [4]   // Chemical Conductivity
        [5]   // Pump pressure
   FALSE : BOOL;   // Always false bit
   FC45_NbCycBeforeMaint : DINT := 899;
   FinalRinseCond : REAL := 34.34375;
   I_Chem_Cond : DINT := 4000;   // Chemical water conductivity
   I_Chm_1_Lvl_Sw : BOOL := 1;   // Chemical Pump #1 level switch
   I_Chm_2_Lvl_Sw : BOOL := 1;   // Chemical Pump #2 level switch
   I_Chm_3_Lvl_Sw : BOOL;   // Chemical Pump #3 level switch
   I_Chm_4_Lvl_Sw : BOOL;   // Chemical Pump #4 level switch
   I_Dry_RTD : DINT := 223;   // Drying RTD
   I_Final_Rinse_Cond : DINT := 9495;   // Final rinse water conductivity
   I_Ld_Dr_Cls_Sw : BOOL := 1;   // Load door close
   I_Ld_Dr_Obs_Sw : BOOL := 1;   // Load door obstruction switch
   I_MCR : BOOL := 1;   // MCR input
   I_Mtr_Ovrld : BOOL;   // Motor overload
   I_Pump_Press : DINT := 12566;   // Recirculation pump pressure
   I_Pure_Water_Filling_Auth : BOOL := 1;
   I_Pw_Tnk_Lvl_Sw : BOOL;   // Pure water tank level switch
   I_Pw_Tnk_RTD : DINT := 214;   // Pure water tank RTD
   I_Pw_Tnk_Sft_Lvl_Sw : BOOL := 1;   // Pure water tank safety level switch
   I_Shlf_Sw : BOOL := 1;   // Shelf switch
   I_Smp_Lvl_Hgh : BOOL;   // Sump high level switch
   I_Smp_Lvl_Lw : BOOL;   // Sump low level switch
   I_Smp_RTD : DINT := 212;   // Sump RTD
   I_Smp_Sft_Lvl_Sw : BOOL := 1;   // Sump safety level switch
   I_Unld_Dr_Cls_Sw : BOOL;   // Unload door close
   I_Unld_Dr_Obs_Sw : BOOL;   // Unload door obstruction switch
   I_UnldDr_ClseSlnce_Bttn : BOOL;   // Door Close/ Silence button Unload Side
   I_UnldDr_Opn_Bttn : BOOL;   // Door Open button Unload side
   iAlarmToSCADA : INT;
   iAuditTrailExportStatus : INT;   // Export Status Of the Audit Trail : 0 - Initial Status Code 200 - Transfer Succesfull
   iDelayBeforeFillingAuthAlarmMM : DINT := 1;
   iDelayBeforeFillingAuthAlarmSS : DINT;
   iInactivityLogoutTime : DINT;   // Inactivity Logout Time In Minutes
   iInactivityPeriod : DINT := 1;   // Inactivity Period before Logout * Value Must be greater than 0
   iPWClosingDelayMM : DINT;
   iPWClosingDelaySS : DINT;
   iSCADACycleCompleteTimeHr : INT := 14;
   iSCADACycleCompleteTimeMin : INT := 16;
   iSCADACycleCompleteTimeSec : INT := 52;
   iSerialModuleActivateDeactivateInhibit : DINT;   // Set Bit 2 Of Word to Inhibited Serial M Reset Bit 2 Of Word to Un-inhibited
   L32E_ETH_Cfg : TIMER := (PRE := 30000);   // Delay for Ethernet port initialization
   Language_English : STRING := 'en-CA';
   LastCheckNbrDays : DINT := 9711;
   LastRecircSumpDrainTemp : REAL := 41.0;
   Load : Doors := (Obstruction := 1, Closed := 1, PreviousScreen := 99, Closing := 1, Delay12S := 12000, Delay1250ms := 1250, Step15 := 1, MsgOpening := 2, MsgClosing := 8, CurrentScreen := 99);
   LoadDoorClosing : BOOL;
   LoadDoorOpening : BOOL;
   MaintainCloseLd : BOOL := 1;
   MaintainCloseUnld : BOOL;
   MaintainOpenLd : BOOL;
   MaintainOpenUnld : BOOL;
   MaintenanceDueDays : DINT := 5;
   MinorFaultBits : DINT := 144;
   msg : BOOL[512];
   Msg_Abort : SINT;
   Msg_CalibChem : SINT;
   Msg_CalibFrinse : SINT;
   Msg_CalibPress : SINT;
   Msg_Door : SINT;   // 1= Door(s) not closed
   Msg_DoorSteps : INT := 8;   // Display Safety Door Test Messages
   Msg_EditCalib : SINT;   // Screen 103 Msg Display
   Msg_Phase : DINT := 19;
   Msg_PwrUp : DINT := 2;
   Msg_Shutdown : SINT;
   Msg_TempSp : SINT;   // HMI Information Message tag
   Msg_TempSp_Ack : BOOL;
   MsgIterator : DINT;   // Iterator to Iterate Through all Printout Mesage
   MsgNumbers : DINT := 246;
   N13 : DINT := 139198;
   Non_Vented_with_Dry_Option : BOOL := 1;
   NonVented_Without_Dry_Option : BOOL;
   NOT_USED : SINT[3] := ([1] := 48, [2] := -13);
        [1]   // Not Used
        [2]   // Not Used
   NumInput : UDT_NUMERIC_INPUT[65] := ([2].value := 1210, [3].value := 14526001, [3].caption := 14526001, [4].value := 2090, [4].caption := 2090, [5].value := 8, [5].caption := 8, [6].value := 14, [6].caption := 14, [7].value := 1, [9].value := 2, [9].caption := 2, [15].value := 10, [16].value := 1, [19].value := 2, [19].caption := 2, [20].value := 8, [20].caption := 8, [21].caption := 9999, [22].value := 10, [23].value := 900, [24].value := 99, [24].caption := 99, [25].value := 90, [25].caption := 90, [26].value := 180, [27].value := 60, [28].value := 10, [28].caption := 10, [29].value := 2026, [30].value := 8, [31].value := 12, [32].value := 13, [33].value := 35, [34].value := 35, [35].value := 6, [35].caption := 6, [38].value := 8, [38].caption := 8, [40].value := 20, [40].caption := 20, [42].value := 9, [42].caption := 9, [44].value := 2, [44].caption := 2, [47].value := 2, [47].caption := 2, [52].value := 20, [52].caption := 20, [53].value := 12, [54].value := 12, [55].value := 12, [56].value := 12, [57].value := 135, [58].value := 135, [59].value := 58, [60].value := 58, [61].value := 12, [62].value := 12, [63].value := 3,
        [64].value := 3);   // Numeric input
        [0]   // NOT USED
        [0].value   // Service Password
        [0].enter   // Service Numeric pad Enter key pressed
        [0].hds   // Handshake
        [10]   // Numeric input min, Sump fill alarm time sec
        [11]   // Drying time in minutes
        [12]   // Drying time in seconds
        [13]   // Not Used
        [14]   // Final rinse time (minutes) numeric input
        [15]   // Final rinse time (seconds) numeric input
        [16]   // Final rinse number of final rinse numeric input
        [17]   // Final rinse minimum number of final rinse numeric input
        [18]   // Final rinse conductivity set point rinse numeric input
        [19]   // Numeric Input On time
        [19].enter   // Numeric input On Time
        [1]   // NOT USED
        [1].enter   // Supervisor Login numeric pad entry
        [20]   // Numeric Input Off time
        [20].enter   // Numeric input Off Time
        [21]   // NOT USED
        [21].enter   // Numeric input to set current Sup. password
        [22]   // Cycle Counter numeric input
        [23]   // NB of cycles before next maintenance numeric input
        [24]   // Calib Chemical Value numeric input
        [25]   // Calib Frinse Value, numeric input
        [26]   // Chemical volume injected, numeric input
        [27]   // Calib Pressure PSI, numeric input
        [28]   // Numeric input, Audible alarm activation time sec.
        [29]   // Set Year numeric input
        [29].value   // Supervisor year entry
        [29].enter   // Supervisor year entry confirmation
        [29].hds   // Supervisor year entry confirmation handshake
        [2]   // Numeric input RTD calibration
        [30]   // Set Month numeric input
        [30].value   // Supervisor month entry
        [30].enter   // Supervisor month entry confirmation
        [30].hds   // Supervisor month entry confirmation handshake
        [31]   // Set Date numeric input
        [31].value   // Supervisor day entry
        [31].enter   // Supervisor day entry confirmation
        [31].hds   // Supervisor day entry confirmation handshake
        [32]   // Set Hour numeric input
        [32].value   // Supervisor hour entry
        [32].enter   // Supervisor hour entry confirmation
        [32].hds   // Supervisor hour entry confirmation handshake
        [33]   // Set Min numeric input
        [33].value   // Supervisor minute entry
        [33].enter   // Supervisor minute entry confirmation
        [33].hds   // Supervisor minute entry confirmation handshake
        [34]   // Set Sec numeric input
        [34].value   // Supervisor second entry
        [34].enter   // Supervisor second entry confirmation
        [34].hds   // Supervisor second entry confirmation handshake
        [35]   // Set Min Max injection Time Cond.
        [35].enter   // Min. Max Injection time cond. numeric pad entry
        [36]   // Set Sec Max injection Time Cond.
        [36].enter   // Sec. Max Injection time cond. numeric pad entry
        [37]   // NOT USED
        [37].enter   // Numeric input to set new Sup. password
        [38]   // Numeric input min, Pure Water Tank fill alarm time min.
        [39]   // Numeric input min, Pure Water Tank fill alarm time sec
        [3]   // Serial Number Numeric Pad entry 8 Last digits
        [3].enter   // Serial Number Numeric pad entry 8 last digits
        [3].hds   // Serial Number Numeric pad entry HDS tag
        [40]   // Numeric input min, Pure Water Tank heating alarm time min.
        [41]   // Numeric input min, Pure Water Tank heating alarm time sec
        [42]   // Numeric input, Maximum number of final rinses
        [43]   // Numeric input sec, Drain extension time
        [44]   // Numeric input min, Vapor removal time min.
        [45]   // Numeric input min, Vapor removal time sec
        [46]   // Numeric input m, Altitude m.
        [47]   // Numeric input min, Drying cooling time min.
        [47].enter   // Numeric Input Drying cooling Time Min
        [48]   // Numeric input min, Drying cooling time sec
        [48].enter   // Numeric Input Drying cooling Time Sec
        [49]   // NOT USED
        [4]   // Numeric input for Year
        [50]   // Numeric Input Recirc. Neutralization Time, Min
        [51]   // Numeric Input Recirc. Neutralization Time, Sec
        [52]   // Numeric input, Heating interval alarm time
        [53]   // PMPack 1 Month Setpoint
        [54]   // PMPack 2 Month Setpoint
        [55]   // PMPack 3 Month Setpoint
        [56]   // PMPack 4 Month Setpoint
        [57]   // PMPack 1 Cycle Count
        [58]   // PMPack 2 Cycle Count
        [59]   // PMPack 3 Cycle Count
        [5]   // Numeric input for Month
        [60]   // PMPack 4 Cycle Count
        [61]   // PMPack 1 Month Accumulation
        [62]   // PMPack 2 Month Accumulation
        [63]   // PMPack 3 Month Accumulation
        [64]   // PMPack 4 Month Accumulation
        [6]   // Numeric input for Date
        [7]   // Numeric input min
        [8]   // Numeric input sec
        [9]   // Numeric input min, Sump fill alarm time min.
   NumInputReal : UDT_NUMERIC_INPUT_REAL[17] := ([0].value := 59.46558, [0].caption := 4.1, [2].value := 65.6, [3].value := 0.5, [3].caption := 0.5, [4].value := 0.8, [4].caption := 80.0, [5].value := 5.0, [5].caption := 5.0, [6].value := 50.0, [7].value := 0.34473723, [7].caption := 0.34473723, [8].value := 18.0, [8].caption := 0.9, [9].value := 1.0, [9].caption := 1.0, [10].value := 1.0, [10].caption := 1.0, [11].value := 1.0, [11].caption := 1.0, [12].value := 1.0, [12].caption := 1.0, [13].value := 234.0, [13].caption := 234.0, [14].value := 226.0, [14].caption := 226.0, [15].value := 1097.0, [15].caption := 1097.0, [16].value := 1084.0, [16].caption := 1084.0);
        [0]   // Pressure Calibration Numeric input
        [10]   // Numeric Input, Chem 2 Neutralization Ratio
        [11]   // Numeric Input, Chem 3 Neutralization Ratio
        [12]   // Numeric Input, Chem 4 Neutralization Ratio
        [1]   // Wash Conductivity Setpint 1st injection
        [2]   // Temperature Sp numeric input PW-W- R
        [3]   // Sump heating rate °C
        [4]   // % Before ON-Off sequence
        [4].enter   // % Bebore On-Off sequence numeric input
        [5]   // Low pressure alarm setpoint
        [6]   // Temperature Sp numeric input Final Rinse
        [7]   // Low pressure alarm setpoint bar
        [8]   // Sump heating rate ° F
        [9]   // Numeric Input, Chem 1 Neutralization Ratio
   ONS_SCADA : INT;
   ONS_WSH64 : SINT := 4;
   PmpPres : REAL := 32.122498;
   PreHeatTime : DINT := 40000;
   PressureUnit : BOOL;   // Pressure Unit 0=PSIG 1=BAR
   previous_s108 : DINT := 99;
   printAlarm : STRING := 'Alarm';
   printAlarmMsg : STRING[50] := ([1] := 'LOAD DOOR DID NOT OPEN', [2] := 'LOAD DOOR DID NOT CLOSE', [3] := 'LOAD DOOR OBSTRUCTED', [4] := 'LOAD DOOR OPEN', [5] := 'UNLOAD DOOR DID NOT OPEN', [6] := 'UNLOAD DOOR DID NOT CLOSE', [7] := 'UNLOAD DOOR OBSTRUCTED', [8] := 'UNLOAD DOOR OPEN', [9] := 'SUMP SAFETY WATER LEVEL REACHED', [10] := 'PURE WATER TANK SAFETY WATER LEVEL REACHED', [11] := 'SUMP TOO LONG TO FILL', [12] := 'SUMP DRAIN TOO LONG', [13] := 'SUMP TOO LONG TOO HEAT', [14] := 'SUMP RTD DEFECTIVE', [15] := 'SUMP TEMPERATURE TOO HIGH', [16] := 'PURE WATER TANK TOO LONG TO FILL', [17] := 'PURE WATER TANK DRAIN TOO LONG', [18] := 'PURE WATER TANK TOO LONG TO HEAT', [19] := 'PURE WATER TANK RTD DEFECTIVE', [20] := 'PURE WATER TANK TEMPERATURE TOO HIGH', [21] := 'PURE WATER TANK FAILED TO DUMP', [22] := 'CHEMICAL CONTAINER 1 EMPTY', [23] := 'CHEMICAL CONTAINER 2 EMPTY', [24] := 'CHEMICAL CONTAINER 3 EMPTY', [25] := 'CHEMICAL CONTAINER 4 EMPTY', [26] := 'DRYING TEMPERATURE NOT REACHED', [27] := 'CHEMICAL INJECTION CONDUCTIVITY SETPOINT NOT REACHED', [28] := 'FINAL RINSE CONDUCTIVITY SETPOINT NOT REACHED', [29] := 'FINAL RINSE CONDUCTIVITY SYSTEM DEFECTIVE', [30] := 'CHEMICAL CONDUCTIVITY SYSTEM DEFECTIVE', [31] := 'PRESSURE TRANSMITTER DEFECTIVE', [32] := 'PUMP PRESSURE TOO LOW', [33] := 'MOTOR OVERLOAD DETECTED', [34] := 'MAINTENANCE DUE', [35] := 'BOTH DOORS OPEN', [36] := 'DRYING RTD DEFECTIVE', [37] := 'MASTER CONTROL RELAY DEACTIVATED', [38] := 'PURE WATER TANK TEMPERATURE ABOVE TEMPERATURE RANGE ALLOWED', [39] := 'PURE WATER TANK TEMPERATURE BELOW TEMPERATURE RANGE ALLOWED', [40] := 'BATTERY LOW', [41] := 'I/O COMMUNICATION HAS BEEN LOST', [42] := 'WAITING FOR PURE WATER FILLING AUTHORIZATION', [43] := 'AUDIT TRAIL LOW STORAGE MEMORY');
   PrintChemCondValue : REAL;
   printEvent : STRING[5] := ([0] := 'CYCLE STOPPED:', [1] := 'CYCLE RESUMED:', [2] := 'CYCLE ABORTED:', [3] := 'MACHINE SERVICE MODE:');
   PrintFrinseCondValue : REAL;
   PrintHardware : STRING[29] := ([0] := '*******  HARDWARE OPTIONS  *******', [1] := 'MODEL: 400XLS', [2] := 'MODEL: 500XLS', [3] := 'NUMBER OF DOOR(S):', [4] := '1', [5] := '2', [6] := 'NON-RECIRCULATED HEATED PURE WATER RINSE SYSTEM:', [7] := 'YES', [8] := 'NO', [9] := 'NON-VENTED VAPOR CONDENSER:', [10] := 'VENTED WITH DRYING SYSTEM:', [11] := 'NON-VENTED WITH DRYING SYSTEM:', [12] := 'HEAT RECOVERY TANK SYSTEM:', [13] := 'PROCESS MONITORING SYSTEM:', [14] := 'DRAIN DISCHARGE COOL DOWN SYSTEM:', [15] := 'ADDITIONAL CHEMICAL PUMPS (PUMP 3 AND PUMP 4):', [16] := 'CONDENSATE RETURN COOL DOWN SYSTEM:', [17] := 'ELECTRICAL HEATED UNIT:', [18] := 'PRINTER OPTION:', [19] := 'CR2 RELAY OPERATING MODE:', [20] := 'CYCLE COMPLETED SIGNAL', [21] := 'EXTERNAL PURE WATER VALVE', [23] := 'Email & SMS Notification ', [25] := 'AUDIT TRAIL:', [26] := 'BATCH REPORT:', [27] := 'CYCLE VALIDATION:', [28] := 'ELECTRONIC SIGNATURE:');
   printID : STRING[6] := ([0] := 'POWER UP :', [1] := 'RELIANCE 400XLS', [2] := 'RELIANCE 500XLS', [3] := 'S/N:', [4] := 'SOFTWARE VERSION', [5] := '13968431 Rev. A');
        [5]   // Software version
   PrintIndex : DINT;
   PrintoutMsgHandshake : BOOL;   // Flag Send to HMI to Acknowledge Reception of Message
   PrintoutMsgNotification : BOOL[512];   // Flag Send by HMI when a Message is sended to PLC
   PrintSystemOption : STRING[29] := ([0] := '*******  SYSTEM OPTIONS  *******', [1] := 'CYCLE COUNTER:', [2] := 'NB OF CYCLES BEFORE NEXT MAINTENANCE:', [3] := 'NEXT MAINTENANCE DATE:', [4] := 'YEAR:', [5] := 'MONTH:', [6] := 'DATE :', [7] := 'SUMP FILL ALARM TIME:', [8] := 'SUMP HEATING INTERVAL ALARM TIME:', [9] := ':', [10] := '0', [11] := '(MIN-SEC)', [12] := 'SEC', [13] := 'PURE WATER TANK FILL ALARM TIME:', [14] := 'PURE WATER TANK HEATING ALARM TIME:', [15] := 'MAXIMUM NUMBRER OF FINAL RINSE:', [16] := 'DRAIN EXTENSION TIME:', [17] := 'VAPOR REMOVAL TIME:', [18] := 'DRYING COOLING TIME:', [19] := 'ALTITUDE:', [20] := 'm', [21] := 'LOW PRESSURE ALARM SETPOINT:', [22] := 'PSIG', [23] := 'bar', [25] := 'INACTIVITY LOGOUT TIME:', [26] := 'MIN', [27] := 'DELAY BEFORE FILLING AUTH ALARM:', [28] := 'PURE WATER CLOSING DELAY:');
   PureWaterTankDrainingDeadLeg : BOOL;
   PureWaterTankFillingRequest : BOOL;
   PureWaterTankTemp : REAL := 21.9;   // Pure water tank temperature
   PWT_DeltaTempNeg : REAL := -8.0;
   PWT_DeltaTempPos : REAL := 8.0;
   Q_Adble_Alrm : BOOL;   // Audible Alarm and /Pilot Light: red connection
   Q_Chm_1 : BOOL;   // Chemical pump #1
   Q_Chm_2 : BOOL;   // Chemical pump #2
   Q_Chm_3 : BOOL;   // Chemical pump #3
   Q_Chm_4 : BOOL;   // Chemical pump #4
   Q_Cld_Wtr_Fll_Vlve : BOOL;   // Cold water sump fill valve
   Q_Cmmn_Alrm : BOOL := 1;   // Dry contact For Alarm
   Q_Cndsr_Hflw_Vlve : BOOL;   // Condenser high flow cold water valve
   Q_Cndsr_Lflw_Vlve : BOOL;   // Condenser low flow cold water valve
   Q_Condensate_Return_Vlve : BOOL;   // Condensate Return CoolDown water valve
   Q_Cyc_Comp : BOOL;   // Dry Contact For Cycle Completed or Pure Water fill valve
   Q_Cyc_Run : BOOL;   // Pilot light: Green connection
   Q_Drn_Cldwn_Vlve : BOOL;   // Drain cool down water valve
   Q_Dry_Fan : BOOL;   // Vapor removal fan / Drying fan
   Q_Dry_Htr : BOOL;   // Drying heating elements
   Q_Dry_Iso_Vlve : BOOL;   // Drying Isolation Valve (Normally Closed Valve)
   Q_Ht_Rcvry_Tnk_Drn_Vlve : BOOL;   // Heat recovery tank drian valve
   Q_Ht_Wtr_Fll_Vlve : BOOL;   // Hot water sump fill valve
   Q_Int_Lght : BOOL := 1;   // Interior Light
   Q_Ld_Dr_Clse_Vlv : BOOL := 1;   // Load door close pilot valve
   Q_Ld_Dr_Opn_Vlv : BOOL;   // Load door open pilot valve
   Q_Pmp_Hgh_Spd : BOOL;   // Pump high speed
   Q_Pmp_Lw_Spd : BOOL;   // Pump low speed
   Q_Pure_Water_Filling_Request : BOOL;   // Pure Water Filling Request
   Q_Pw_Fll_Vlve : BOOL;   // Pure water sump/ Tank fill valve
   Q_Pw_Otlt_Vlve : BOOL := 1;   // Pure water tank outlet valve
   Q_Pw_Tnk_Stm_Vlve : BOOL;   // PWT Steam Valve / Electric Heater
   Q_Smp_drn_Vlve : BOOL := 1;   // Sump drain valve (Normally open valve)
   Q_Smp_Stm_Vlve : BOOL;   // Sump steam valve/ Electrical Heater
   Q_Trsfr_Vlve : BOOL;   // Transfer Valve (Normally Open Valve)
   Q_Unld_Dr_Clse_Vlve : BOOL;   // Unload door close pilot valve
   Q_Unld_Dr_Opn_Vlve : BOOL;   // Unload door open pilot valve
   RcvryWtrTemp : DINT := 41;
   RD_CHASSIS_1 : MESSAGE;
        MessageParameters(ServiceCode := 16#000e, DestinationTag := Chassis_Size_Ret[1], ...)
   RD_CHASSIS_2 : MESSAGE;
        MessageParameters(ServiceCode := 16#000e, DestinationTag := Chassis_Size_Ret[2], ...)
   RecallSafetyCheck : BOOL;
   RemoteDayOfMonth : DINT := 14;   // HMI Date Day
   RemoteDisplayNumber : DINT;   // HMI connection
   RemoteHour : DINT := 10;   // HMI Time Hour
   RemoteMinute : DINT := 31;   // HMI Time Minute
   RemoteMonth : DINT := 8;   // HMI Date Month
   RemoteSecond : DINT := 20;   // HMI Time Second
   RemoteSetDateTime : BOOL := 1;   // HMI Set Date and Time
   RemoteYear : DINT := 2026;   // HMI Date Year
   rSCADACompensatedSetPoint : REAL := 11.417221;
   s007 : DINT := 7;
   sBatchReportCSVName : STRING := '-BATCH_REPORT.csv';
   sBatchReportFolderPath : STRING := '\Storage Card2\CycleReport\';
   sChangeLanguage : STRING := 'en-CA';   // jplv09
   Screen_Ctrl : DINT;   // PLC Screen Request
   sCycleAccepted : STRING := 'CYCLE WAS ACCEPTED BY:';   // Cycle Accepted
   sCycleCounter : STRING := '60';
   sCycleForFileName : STRING := 'CYCLE_';
   sCycleRejected : STRING := 'CYCLE WAS REJECTED BY:';   // Cycle Rejected
   sDate : STRING := '17-08-2026';   // String current date
   sDateTime : STRING := '17-08-2026  -  11:01:29';   // String Date Time
   SelChemi_Remote : SINT;
   SelChemical_Ind : SINT;
   SelChemical_Value : SINT := 3;
   SelChemNeutralizer : UDT_SELECTOR[5];
        [1]   // Chem 1 Neutralizant pump
        [2]   // Chem 2 Neutralizant pump
        [3]   // Chem 3 Neutralizant pump
        [4]   // Chem 4 Neutralizant pump
   SelChemNeutralizerESign : UDT_SELECTOR[5];
   Selector : UDT_SELECTOR[25] := ([0].Value := 1, [1].Indicator := 1, [1].Remote := 1, [2].Value := 1, [2].Indicator := 1, [5].Value := 2, [5].Indicator := 2, [7].Indicator := 1, [8].Value := 3, [10].Value := 3, [14].Value := 1, [14].Indicator := 1, [18].Value := 1, [18].Indicator := 1, [19].Value := 1, [19].Indicator := 1, [22].Value := 1, [23].Value := 2);   // Piloted list selector
        [0]   // Pre-wash modification (treatment selection)
        [0].Value   // Pre-wash's selector list indicator
        [0].Indicator   // Pre-wash's selector list indicator
        [0].Remote   // Pre-wash's selector list remote control tag
        [14]   // Drying mode piloted list selector
        [15]   // Drying temperature (Celsius) piloted list selector
        [16]   // Drying temperature (Fahrenheit) piloted list selector
        [17]   // Heat sensitive drying parameter
        [18]   // Final rinse heating piloted list selector
        [19]   // Final rinse drained piloted list selector
        [1]   // Pre-wash modification (heating selection)
        [1].Value   // Pre-wash's heating selector list value
        [1].Indicator   // Pre-wash's heating selector list indicator
        [1].Remote   // Pre-wash's heating selector list remote control tag
        [20]   // Final rinse recirculated piloted list selector
        [21]   // Final rinse type piloted list selector
        [22]   // Rinse Treatment selector
        [23]   // Audible alarm op. mode selector
        [2]   // Pre-wash modification (water port selection)
        [2].Remote   // Pre-wash's water port selector list remote control tag
   SelectorView : UDT_SELECTOR[3];   // Piloted list selector for cycle view menu
        [0]   // Pre-wash view (treatment selection)
        [0].Value   // Pre-wash's selector list indicator
        [0].Indicator   // Pre-wash's selector list indicator
        [0].Remote   // Pre-wash's selector list remote control tag
        [1]   // Wash view (treatment selection)
        [1].Value   // Pre-wash's heating selector list value
        [1].Indicator   // Pre-wash's heating selector list indicator
        [1].Remote   // Pre-wash's heating selector list remote control tag
        [2]   // Rinse view (treatment selection)
        [2].Remote   // Pre-wash's water port selector list remote control tag
   Set_ConfigControl : DINT;
   Set_TCP_Config : UDT_TCPSetAllConfig := (IPAddress := 16#c0a8_0101, SunbNetMask := 16#ffff_ff00);
   sHyphen : STRING := '-';
   SimGenEnabled : BOOL;   // SimGen enable bit 1= Simgen ON
   sNullCharacters : STRING;   // Empty String
   SPV_19 : BOOL := 1;   // Screen 80 Enabled/Disabled Pump pressure monitoring
   sTime : STRING := '11:01:29';   // String current time
   StringInput : UDT_STRING_INPUT[6] := ([0].Value := 'STERIS', [0].Caption := '1', [1].Value := 'CIP 100', [1].Caption := 'CIP 100', [2].Value := 'CIP 200', [2].Caption := 'CIP 200', [3].Value := 'Pump 3', [3].Caption := 'N/A', [4].Value := 'Pump 4', [4].Caption := 'N/A');
        [0].Enter   // Screen 99 ASCII pad Change Cycle Name
        [1]   // Chemical 1 Name
   SumpAlarmFillTime : DINT := 120000;
   SumpHeatAlmRate : REAL := 1.0;
   SumpTemp : REAL := 21.7;   // Sump temperature in °C
   SumpTempToCool : REAL := 41.0;   // Sump temperature in °C
   sUnderscore : STRING := '_';
   tAuditTrailRemoteClearHistory : TIMER := (PRE := 2000);
   tDelayBeforeFillingAuthAlarm : TIMER := (PRE := 60000);
   tDelayBeforeTankFillingAuthAlarm : TIMER := (PRE := 60000);
   TempUnit : BOOL;   // Temperature Units 0= Celcius 1 = Farhenheit
   Tpb : DINT[11] := ([5] := 8, [7] := 4096, [10] := 63983);
        [0].0   // DOOR button Ready Mode screen Cycle complete screen Manual Injection screen
        [0].1   // Close Door (load door button) Door Init.screen
        [0].10   // HMI Chemical Pump 1 button
        [0].11   // HMI Chemical Pump 2 button
        [0].12   // HMI Chemical Pump 3 button
        [0].13   // HMI Chemical Pump 4 button
        [0].14   // HMI Service Mode Open Pilot Valve button
        [0].15   // HMI Service Mode Stop Load Door button
        [0].16   // HMI Service Mode Open Pilot Valve Unload Door button
        [0].17   // HMI Service Mode Stop Unload Door button
        [0].18   // HMI Transfer Valve
        [0].19   // HMI Sump Heating
        [0].2   // Close Door (Unload door button) Door Init.screen
        [0].20   // HMI Pure Water Outlet Valve
        [0].21   // HMI Pure Water Tank Heating
        [0].22   // HMI Sump Cold Water Fill Valve
        [0].23   // HMI Cool-Down Valve
        [0].24   // HMI Cold Water Fill Valve
        [0].25   // HMI Sump Drain Valve
        [0].26   // HMI Pure Water Fill Valve
        [0].27   // HMI Heat Recovery Drain Valve
        [0].28   // HMI Condenser Low Flow Valve
        [0].29   // HMI Condenser Low Flow Valve
        [0].3   // HMI CYCLE START button
        [0].30   // HMI Drying Fan Button
        [0].31   // HMI Drying Element Button
        [0].4   // HMI STOP CYLE Button
        [0].5   // HMI RESUME button
        [0].6   // HMI Start Pump Low speed button
        [0].7   // HMI Start Pump High speed button
        [0].8   // Screen 18 HMI Print Cycle Parameters button
        [0].9   // Exit Service Mode button
        [10].0   // PMPack 1 Enable Bit
        [10].1   // PMPack 2 Enable Bit
        [10].11   // Service Mode Entered Email Enable
        [10].12   // Superviser Mode Entered Email Enable
        [10].13   // Not Used
        [10].14   // Preventive Maintenance Due Email Enable
        [10].15   // Process Alarms Email Enable
        [10].16   // Pure Water Filling Request
        [10].2   // PMPack 3 Enable Bit
        [10].3   // PMPack 4 Enable Bit
        [10].4   // PMPack Cycle Count
        [10].5   // Cycle Started Email Enable
        [10].6   // Cycle Completed Email Enable
        [10].7   // Cycle Aborted Email Enable
        [10].8   // Cycle Values Changed Email Enable
        [1]   // Not Used pB
        [1].0   // HMI Isolation Valve button
        [1].1   // HMI Service Mode Close Pilot Valve Unload Door button
        [1].10   // HMI Service Mode Navigation
        [1].11   // HMI Service Mode Navigation
        [1].12   // HMI Service Mode Navigation
        [1].13   // HMI Service Mode Navigation
        [1].14   // HMI Service Mode Navigation
        [1].15   // HMI Service Mode Navigation
        [1].16   // HMI Service Mode Navigation
        [1].17   // HMI Service Mode Navigation
        [1].18   // HMI Service Mode Navigation
        [1].19   // HMI Service Mode Navigation
        [1].2   // HMI Cycle Run Pilot Valve
        [1].20   // HMI Service Mode Navigation
        [1].21   // HMI Service Mode Navigation
        [1].22   // HMI Service Mode Navigation
        [1].23   // HMI Service Mode Navigation
        [1].24   // HMI Service Mode Navigation
        [1].25   // HMI Service Mode Navigation
        [1].26   // HMI Service Mode Navigation
        [1].27   // HMI Service Mode Navigation
        [1].28   // HMI Service Mode Navigation
        [1].29   // HMI Service Mode Navigation
        [1].3   // HMI Dry Contact For Alarm
        [1].30   // HMI Service Mode Navigation
        [1].31   // HMI Service Mode Navigation
        [1].4   // Hmi Interior Light
        [1].5   // HMI Dry Contact for Cycle Completed
        [1].6   // HMI Audible Alarm/Red Status Light/Alarm Signal Relay
        [1].7   // HMI Service Mode Navigation
        [1].8   // HMI Service Mode Navigation
        [1].9   // HMI Service Mode Navigation
        [2].0   // HMI Navigation (Service Mode)
        [2].1   // HMI Navigation (Service Mode)
        [2].10   // Next page
        [2].11   // Previous page
        [2].12   // Exit button
        [2].13   // Exit button
        [2].14   // HMI Navigation (Operator Mode)
        [2].15   // HMI Navigation (Operator Mode)
        [2].16   // Manual injection resume cycle button
        [2].17   // HMI Mute Button
        [2].18   // Screen 31 Change Cycle set-up button
        [2].19   // Screen 35, 36, 37 X button
        [2].2   // HMI Navigation (Service Mode)
        [2].20   // Screen 35 Next button
        [2].21   // Screen 36 Previous button
        [2].22   // Screen 36 Next button
        [2].23   // Screen 37 Previous button
        [2].24   // EXTRACare button
        [2].25   // ENVIROCare button
        [2].26   // PLASTIC button
        [2].27   // STANDARD button
        [2].28   // RINSECare button
        [2].29   // DESCALER button
        [2].3   // Screen 31 Exit button
        [2].30   // CYCLE 6 button
        [2].31   // CYCLE 7 button
        [2].4   // Calibration Start/Stop button
        [2].5   // Done Entering Data
        [2].6   // Restore default value
        [2].7   // Calibration button
        [2].8   // Exit button
        [2].9   // Sump RTD calibration button
        [3].0   // CYCLE 8 button
        [3].1   // CYCLE 10 button
        [3].10   // Screen 39 Drying button
        [3].11   // HMI Nav. (Sup. mode) X Button Pw-W-R, FR, Drying conf. screens
        [3].12   // Extra Care button
        [3].13   // Enviro Care button
        [3].14   // Plastic Care button
        [3].15   // Standard button
        [3].16   // Rinse care button
        [3].17   // Descaler button
        [3].18   // Cycle 7 button
        [3].19   // Cycle 8 button
        [3].2   // CYCLE 11 button
        [3].20   // Cycle 9 button
        [3].21   // Cycle 10 button
        [3].22   // Cycle 11 button
        [3].23   // Exit to ready screen
        [3].24   // HMI navigation
        [3].25   // HMI navigation
        [3].26   // HMI navigation
        [3].27   // HMI navigation
        [3].28   // HMI navigation
        [3].29   // HMI Abort button
        [3].3   // Screen 38 X button
        [3].30   // HMI YES button (Abort screen)
        [3].31   // HMI NO button (Abort screen)
        [3].4   // Screen 38 Parameters button
        [3].5   // Screen 39 X button
        [3].6   // HMI Nav. (Sup. mode) Pre-wash selection
        [3].7   // Screen 39 Wash button
        [3].8   // Screen 39 Rinse button
        [3].9   // Screen 39 Final Rinse button
        [4].0   // HMI Nav. (Sup. mode) Save Button pre-wash screen
        [4].1   // Factory Reset Request
        [4].11   // Save button Final Rinse screen
        [4].12   // Wake button of the shutdown screen
        [4].13   // Shutdown button of the ready mode screen
        [4].14   // Drying RTD calibration button
        [4].15   // Pure water tank RTD calibration button
        [4].16   // Exit button (readymode screen)
        [4].17   // Goto option screen
        [4].18   // HMI Nav. (Sup. mode) Save Button Rinse screen
        [4].19   // HMI Next Ready Mode Screen
        [4].2   // HMI Nav. Next screen (screen 41)
        [4].20   // HMI Previous Ready Mode Screen
        [4].21   // HMI View Cycle general data
        [4].22   // HMI View Pre-Wash data
        [4].23   // HMI View Wash data
        [4].24   // HMI View Wash data 2
        [4].25   // HMI View Wash data 3
        [4].26   // HMI View Rinse data
        [4].27   // HMI View Final Rinse data
        [4].28   // HMI View Final Rinse data 2
        [4].29   // HMI View Drying data
        [4].3   // X button Chemical pump sel 2nd injection screen 92
        [4].30   // HMI Condensate Return Valve
        [4].31   // HMI Exit View cycle mode
        [4].4   // HMI Nav. Next screen button Wash 2 screen 42
        [4].5   // Save button Chemical 2nd Injection screen 92
        [4].6   // Save button Drying screen
        [5].0   // Screen 64 HMI Service Mode Close Pilot Valve button
        [5].1   // HMI Select cycle pump speed (Sup. Mode)
        [5].10   // Exit button to supervisor 2 screen
        [5].11   // Display Set date screen
        [5].12   // Previous to supervisor screen button
        [5].13   // Display Set time screen
        [5].2   // HMI Select cycle water level (Sup. Mode)
        [5].24   // Screen 33 Chemical Pumps (calibration)
        [5].25   // Screen 54 START button
        [5].26   // Screen 54 X button
        [5].27   // Screen 54 Print button
        [5].3   // HMI Select cycle permission (lock/unlock) (Sup. Mode)
        [6].1   // Display Water Port Screen (56)
        [6].10   // X button Cond. Sp screen 91
        [6].11   // Concentration button 2nd injection screen 43
        [6].12   // X button Concentration screen 90
        [6].13   // Save button Water Port screen 56
        [6].14   // Save button Heating screen 57
        [6].15   // Save button Time Min Sec screen 58
        [6].16   // X button Inj Type screen screen 60
        [6].17   // Water Port button Rinse Screen (48)
        [6].18   // HMI Nav. Rinse Heating button
        [6].19   // HMI Nav. Time button Rinse screen 48
        [6].2   // HMI Nav. (Sup. mode) Heating button
        [6].20   // Treatment selection screen Screen 39 Reset to default button
        [6].21   // YES button Reset to Default Cycles Values Screen 93
        [6].22   // No button Reset to Default Cycles Values Screen 93
        [6].3   // HMI Nav. Time button Wash screen
        [6].31   // Screen 1 Monitoring option is present NO button
        [6].4   // Water Port button Pre-Wash Screen (40)
        [6].5   // HMI Nav. Prewash screen Heating button
        [6].6   // HMI Nav. Time button Prewashscreen
        [6].7   // X button Water Port Screen (56)
        [6].8   // X button Temperature Screen 57
        [6].9   // X button Time Min Sec 58
        [7].0   // HMI Nav. Chemical button screen 59
        [7].1   // Inj. Type button screen 42
        [7].10   // Non-Vented Vapor Condenser
        [7].11   // Vented with drying system
        [7].12   // Non-Vented with Drying system
        [7].2   // Concentration button 1st injection screen 42
        [7].22   // Screen 38 Next screen button
        [7].23   // Screen 99 Previous screen button
        [7].24   // Screen 99 X button
        [7].25   // Screen 100 No Button
        [7].26   // Screen 101 Cancel Button
        [7].27   // Screen 101 Door Test Open Load Door button
        [7].29   // Screen 101 Door Test Open Load Door button
        [7].3   // Conductivity Sp button screen 42
        [7].30   // Screen 101 Door Test Close Load Door button
        [7].31   // Screen 1 Monitoring option is present YES button
        [7].4   // Chemical button 2nd injection screen 43
        [7].5   // Save button Chemical 1st Injection screen 59
        [7].6   // X button Chemical selectiuon 1st injection screen 59
        [7].7   // Save button Inj. Type 1 st Injection screen 60
        [7].8   // Save button Concentration screen 90
        [7].9   // Save button Cond Sp screen 91
        [8].0   // Screen 31 Chemical Parameters button
        [8].1   // X button
        [8].10   // Screen 49 Next screen button
        [8].11   // Screen 80 Previous screen button
        [8].12   // Screen 80 Neutralization parameters button
        [8].13   // Screen 81, 82 X Button
        [8].14   // Screen 81 Next screen button
        [8].15   // Screen 81 Previous screen button
        [8].16   // Screen 80 Audible alarm mode button
        [8].17   // Screen 83 Previous screen button
        [8].18   // Screen 30 Automatic Shutdown button 1= Yes 0 = No
        [8].19   // Screen 32 Edit Calibration button
        [8].2   // Screen 94 Next screen button
        [8].20   // Screen 102 X button
        [8].21   // Screen 102 Print Calibration button
        [8].22   // Screen 103 OK Button
        [8].23   // Screen 103 X button
        [8].24   // Screen 102 Sump RTD button
        [8].25   // Screen 102 PWT RTD button
        [8].26   // Screen 102 Dry RTD button
        [8].27   // Screen 102 Pressure button
        [8].28   // Screen 102 Chemical button
        [8].29   // Screen 102 Final Rinse button
        [8].3   // Screen 95 Previous screen button
        [8].30   // Screen 88 Print Hardware options button
        [8].31   // Screen 79 Print System options button
        [8].4   // Screen 95 next screen button
        [8].5   // Screen 96 Previous screen button
        [8].6   // Screen 49 Change password button
        [8].7   // Screen 97 X button
        [8].8   // Screen 31 Units button
        [8].9   // Screen 98 X button
        [9].0   // Ready Mode Screen 18 Process screen button
        [9].1   // Analog screen (30) Process button
        [9].2   // Screen 85 INIT. AENT button
        [9].3   // Screen 10 Next screen button
        [9].4   // PID screen 10, 6, 104 X button
        [9].5   // Screen 6 or 104 Previous screen button
        [9].6   // Screen 84 X or CANCEL button
   TpbImage : DINT[11] := ([5] := 8, [7] := 4096, [10] := 63983);
        [0].0   // DOOR button Ready Mode screen Cycle complete screen Manual Injection screen
        [0].1   // Close Door (load door button) Door Init.screen
        [0].10   // HMI Chemical Pump 1 button
        [0].11   // HMI Chemical Pump 2 button
        [0].12   // HMI Chemical Pump 3 button
        [0].13   // HMI Chemical Pump 4 button
        [0].14   // HMI Service Mode Open Pilot Valve button
        [0].15   // HMI Service Mode Stop Load Door button
        [0].16   // HMI Service Mode Open Pilot Valve Unload Door button
        [0].17   // HMI Service Mode Stop Unload Door button
        [0].18   // HMI Transfer Valve
        [0].19   // HMI Sump Heating
        [0].2   // Close Door (Unload door button) Door Init.screen
        [0].20   // HMI Pure Water Outlet Valve
        [0].21   // HMI Pure Water Tank Heating
        [0].22   // HMI Sump Cold Water Fill Valve
        [0].23   // HMI Cool-Down Valve
        [0].24   // HMI Cold Water Fill Valve
        [0].25   // HMI Sump Drain Valve
        [0].26   // HMI Pure Water Fill Valve
        [0].27   // HMI Heat Recovery Drain Valve
        [0].28   // HMI Condenser Low Flow Valve
        [0].29   // HMI Condenser Low Flow Valve
        [0].3   // HMI CYCLE START button
        [0].30   // HMI Drying Fan Button
        [0].31   // HMI Drying Element Button
        [0].4   // HMI STOP CYLE Button
        [0].5   // HMI RESUME button
        [0].6   // HMI Start Pump Low speed button
        [0].7   // HMI Start Pump High speed button
        [0].8   // Screen 18 HMI Print Cycle Parameters button
        [0].9   // Exit Service Mode button
        [1]   // Not Used pB
        [1].0   // HMI Isolation Valve button
        [1].1   // HMI Service Mode Close Pilot Valve Unload Door button
        [1].10   // HMI Service Mode Navigation
        [1].11   // HMI Service Mode Navigation
        [1].12   // HMI Service Mode Navigation
        [1].13   // HMI Service Mode Navigation
        [1].14   // HMI Service Mode Navigation
        [1].15   // HMI Service Mode Navigation
        [1].16   // HMI Service Mode Navigation
        [1].17   // HMI Service Mode Navigation
        [1].18   // HMI Service Mode Navigation
        [1].19   // HMI Service Mode Navigation
        [1].2   // HMI Cycle Run Pilot Valve
        [1].20   // HMI Service Mode Navigation
        [1].21   // HMI Service Mode Navigation
        [1].22   // HMI Service Mode Navigation
        [1].23   // HMI Service Mode Navigation
        [1].24   // HMI Service Mode Navigation
        [1].25   // HMI Service Mode Navigation
        [1].26   // HMI Service Mode Navigation
        [1].27   // HMI Service Mode Navigation
        [1].28   // HMI Service Mode Navigation
        [1].29   // HMI Service Mode Navigation
        [1].3   // HMI Dry Contact For Alarm
        [1].30   // HMI Service Mode Navigation
        [1].31   // HMI Service Mode Navigation
        [1].4   // Hmi Interior Light
        [1].5   // HMI Dry Contact for Cycle Completed
        [1].6   // HMI Audible Alarm/Red Status Light/Alarm Signal Relay
        [1].7   // HMI Service Mode Navigation
        [1].8   // HMI Service Mode Navigation
        [1].9   // HMI Service Mode Navigation
        [2].0   // HMI Navigation (Service Mode)
        [2].1   // HMI Navigation (Service Mode)
        [2].10   // Next page
        [2].11   // Previous page
        [2].12   // Exit button
        [2].13   // Exit button
        [2].14   // HMI Navigation (Operator Mode)
        [2].15   // HMI Navigation (Operator Mode)
        [2].16   // Manual injection resume cycle button
        [2].17   // HMI Mute Button
        [2].18   // Screen 31 Change Cycle set-up button
        [2].19   // Screen 35, 36, 37 X button
        [2].2   // HMI Navigation (Service Mode)
        [2].20   // Screen 35 Next button
        [2].21   // Screen 36 Previous button
        [2].22   // Screen 36 Next button
        [2].23   // Screen 37 Previous button
        [2].24   // EXTRACare button
        [2].25   // ENVIROCare button
        [2].26   // PLASTIC button
        [2].27   // STANDARD button
        [2].28   // RINSECare button
        [2].29   // DESCALER button
        [2].3   // Screen 31 Exit button
        [2].30   // CYCLE 6 button
        [2].31   // CYCLE 7 button
        [2].4   // Calibration Start/Stop button
        [2].5   // Done Entering Data
        [2].6   // Restore default value
        [2].7   // Calibration button
        [2].8   // Exit button
        [2].9   // Sump RTD calibration button
        [3].0   // CYCLE 8 button
        [3].1   // CYCLE 10 button
        [3].10   // Screen 39 Drying button
        [3].11   // HMI Nav. (Sup. mode) X Button Pw-W-R, FR, Drying conf. screens
        [3].12   // Extra Care button
        [3].13   // Enviro Care button
        [3].14   // Plastic Care button
        [3].15   // Standard button
        [3].16   // Rinse care button
        [3].17   // Descaler button
        [3].18   // Cycle 7 button
        [3].19   // Cycle 8 button
        [3].2   // CYCLE 11 button
        [3].20   // Cycle 9 button
        [3].21   // Cycle 10 button
        [3].22   // Cycle 11 button
        [3].23   // Exit to ready screen
        [3].24   // HMI navigation
        [3].25   // HMI navigation
        [3].26   // HMI navigation
        [3].27   // HMI navigation
        [3].28   // HMI navigation
        [3].29   // HMI Abort button
        [3].3   // Screen 38 X button
        [3].30   // HMI YES button (Abort screen)
        [3].31   // HMI NO button (Abort screen)
        [3].4   // Screen 38 Parameters button
        [3].5   // Screen 39 X button
        [3].6   // HMI Nav. (Sup. mode) Pre-wash selection
        [3].7   // Screen 39 Wash button
        [3].8   // Screen 39 Rinse button
        [3].9   // Screen 39 Final Rinse button
        [4].0   // HMI Nav. (Sup. mode) Save Button pre-wash screen
        [4].1   // Screen 84 Init. AENT
        [4].11   // Save button Final Rinse screen
        [4].12   // Wake button of the shutdown screen
        [4].13   // Shutdown button of the ready mode screen
        [4].14   // Drying RTD calibration button
        [4].15   // Pure water tank RTD calibration button
        [4].16   // Exit button (readymode screen)
        [4].17   // Goto option screen
        [4].18   // HMI Nav. (Sup. mode) Save Button Rinse screen
        [4].19   // HMI Next Ready Mode Screen
        [4].2   // HMI Nav. Next screen (screen 41)
        [4].20   // HMI Previous Ready Mode Screen
        [4].21   // HMI View Cycle general data
        [4].22   // HMI View Pre-Wash data
        [4].23   // HMI View Wash data
        [4].24   // HMI View Wash data 2
        [4].25   // HMI View Wash data 3
        [4].26   // HMI View Rinse data
        [4].27   // HMI View Final Rinse data
        [4].28   // HMI View Final Rinse data 2
        [4].29   // HMI View Drying data
        [4].3   // X button Chemical pump sel 2nd injection screen 92
        [4].30   // HMI Condensate Return Valve
        [4].31   // HMI Exit View cycle mode
        [4].4   // HMI Nav. Next screen button Wash 2 screen 42
        [4].5   // Save button Chemical 2nd Injection screen 92
        [4].6   // Save button Drying screen
        [5].0   // Screen 64 HMI Service Mode Close Pilot Valve button
        [5].1   // HMI Select cycle pump speed (Sup. Mode)
        [5].10   // Exit button to supervisor 2 screen
        [5].11   // Display Set date screen
        [5].12   // Previous to supervisor screen button
        [5].13   // Display Set time screen
        [5].2   // HMI Select cycle water level (Sup. Mode)
        [5].24   // Screen 33 Chemical Pumps (calibration)
        [5].25   // Screen 54 START button
        [5].26   // Screen 54 X button
        [5].27   // Screen 54 Print button
        [5].3   // HMI Select cycle permission (lock/unlock) (Sup. Mode)
        [6].1   // Display Water Port Screen (56)
        [6].10   // X button Cond. Sp screen 91
        [6].11   // Concentration button 2nd injection screen 43
        [6].12   // X button Concentration screen 90
        [6].13   // Save button Water Port screen 56
        [6].14   // Save button Heating screen 57
        [6].15   // Save button Time Min Sec screen 58
        [6].16   // X button Inj Type screen screen 60
        [6].17   // Water Port button Rinse Screen (48)
        [6].18   // HMI Nav. Rinse Heating button
        [6].19   // HMI Nav. Time button Rinse screen 48
        [6].2   // HMI Nav. (Sup. mode) Heating button
        [6].20   // Treatment selection screen Screen 39 Reset to default button
        [6].21   // YES button Reset to Default Cycles Values Screen 93
        [6].22   // No button Reset to Default Cycles Values Screen 93
        [6].3   // HMI Nav. Time button Wash screen
        [6].31   // Screen 1 Monitoring option is present NO button
        [6].4   // Water Port button Pre-Wash Screen (40)
        [6].5   // HMI Nav. Prewash screen Heating button
        [6].6   // HMI Nav. Time button Prewashscreen
        [6].7   // X button Water Port Screen (56)
        [6].8   // X button Temperature Screen 57
        [6].9   // X button Time Min Sec 58
        [7].0   // HMI Nav. Chemical button screen 59
        [7].1   // Inj. Type button screen 42
        [7].10   // Non-Vented Vapor Condenser
        [7].11   // Vented with drying system
        [7].12   // Non-Vented with Drying system
        [7].2   // Concentration button 1st injection screen 42
        [7].22   // Screen 38 Next screen button
        [7].23   // Screen 99 Previous screen button
        [7].24   // Screen 99 X button
        [7].25   // Screen 100 No Button
        [7].26   // Screen 101 Cancel Button
        [7].27   // Screen 101 Door Test Open Load Door button
        [7].28   // Screen 101 Door Test Close Load Door
        [7].29   // Screen 101 Door Test Open Load Door button
        [7].3   // Conductivity Sp button screen 42
        [7].30   // Screen 101 Door Test Close Load Door button
        [7].31   // Screen 1 Monitoring option is present YES button
        [7].4   // Chemical button 2nd injection screen 43
        [7].5   // Save button Chemical 1st Injection screen 59
        [7].6   // X button Chemical selectiuon 1st injection screen 59
        [7].7   // Save button Inj. Type 1 st Injection screen 60
        [7].8   // Save button Concentration screen 90
        [7].9   // Save button Cond Sp screen 91
        [8].0   // Screen 31 Chemical Parameters button
        [8].1   // X button
        [8].10   // Screen 49 Next screen button
        [8].11   // Screen 80 Previous screen button
        [8].12   // Screen 80 Neutralization parameters button
        [8].13   // Screen 81, 82 X Button
        [8].14   // Screen 81 Next screen button
        [8].15   // Screen 81 Previous screen button
        [8].16   // Screen 80 Audible alarm mode button
        [8].17   // Screen 83 Previous screen button
        [8].18   // Screen 30 Automatic Shutdown button 1= Yes 0 = No
        [8].19   // Screen 32 Edit Calibration button
        [8].2   // Screen 94 Next screen button
        [8].20   // Screen 102 X button
        [8].21   // Screen 102 Print Calibration button
        [8].22   // Screen 103 OK Button
        [8].23   // Screen 103 X button
        [8].24   // Screen 102 Sump RTD button
        [8].25   // Screen 102 PWT RTD button
        [8].26   // Screen 102 Dry RTD button
        [8].27   // Screen 102 Pressure button
        [8].28   // Screen 102 Chemical button
        [8].29   // Screen 102 Final Rinse button
        [8].3   // Screen 95 Previous screen button
        [8].30   // Screen 88 Print Hardware options button
        [8].31   // Screen 79 Print System options button
        [8].4   // Screen 95 next screen button
        [8].5   // Screen 96 Previous screen button
        [8].6   // Screen 49 Change password button
        [8].7   // Screen 97 X button
        [8].8   // Screen 31 Units button
        [8].9   // Screen 98 X button
        [9].0   // Ready Mode Screen 18 Process screen button
        [9].1   // Analog screen (30) Process button
        [9].2   // Screen 85 INIT. AENT button
        [9].3   // Screen 10 Next screen button
        [9].4   // PID screen 10, 6, 104 X button
        [9].5   // Screen 6 or 104 Previous screen button
        [9].6   // Screen 84 X or CANCEL button
   tPureWaterTankClosingDelay : TIMER;
   tPWClosingDelay : TIMER;
   TreatmentPtr : DINT;
   TRUE : BOOL := 1;   // Always true bit
   tStringCopyDebounce : TIMER := (PRE := 1000);
   udtAudibleAlarmMode : UDT_SELECTOR := (Value := 2);
   udtAuditTrail : UDT_AuditTrail;
   udtCSVDataLogBatchReport : UDT_CSVDataLog := (sFileLocation := '\Storage Card2\CycleReport\2026_08_14_13_52_02-CYCLE_60-BATCH_REPORT.csv', sString01 := 'DOOR OPENED:14:17:14');
   udtCSVExport : UDT_CSVExport := (sFileLabel := 'CYCLE_60');
   udtFRHeatingSel : UDT_SELECTOR := (Value := 1, Indicator := 1);
   udtFRLastRinseDrained : UDT_SELECTOR := (Value := 1, Indicator := 1);
   udtFRRecirculation : UDT_SELECTOR;
   udtFRType : UDT_SELECTOR;
   udtPureWaterHandshakeFromSCADA : UDT_PORT_HANDSHAKE_FROM_SCADA;
   udtPureWaterHandshakeToSCADA : UDT_PORT_HANDSHAKE_TO_SCADA;
   Unit : Hrdwre := (Model := 1, PreWtrTnk := 1, Dry := 1, CoolDown := 1, NbChmPmp := 2, Condenser := 1, CWInlet := 1, Printer := 1, AuditTrail := 1, BatchReport := 1);   // Unit Configuration
   UnLoad : Doors := (PreviousScreen := 99, Delay12S := 12000, Delay1250ms := 1250, MsgOpening := 10, MsgClosing := 16, CurrentScreen := 99);
   UnloadDoorClosing : BOOL;
   UnloadDoorOpening : BOOL;
   Valid_Ch_Sizes : DINT[3] := ([0] := 1, [1] := 10, [2] := 11);
   Vented_with_Dry_Option : BOOL;
   WR_CHASSIS_10 : MESSAGE;
        MessageParameters(ServiceCode := 16#0010, LocalElement := Valid_Ch_Sizes[1], ...)
   WR_CHASSIS_11 : MESSAGE;
        MessageParameters(ServiceCode := 16#0010, LocalElement := Valid_Ch_Sizes[2], ...)
END_VAR
